TYPE "UDT_Conv_MultiControl_Status"
VERSION : 0.1
   STRUCT
      OL_Maintenance_Mode : Bool;   // Maintenance mode on
      ER_PE1_Blockage : Bool;   // PE1 blockage
      ER_PE2_Blockage : Bool;   // PE2 blockage
      ER_Motor_1_Fault : Bool;   // Motor has error
      ER_Motor_2_Fault : Bool;   // Motor has error
      ER_Motor_3_Fault : Bool;   // Motor has error
      ER_Motor_4_Fault : Bool;   // Motor has error
      ER_Motor_5_Fault : Bool;   // Motor has error
      ER_Motor_6_Fault : Bool;   // Motor has error
      ER_Motor_7_Fault : Bool;   // Motor has error
      ER_Motor_8_Fault : Bool;   // Motor has error
      ER_Motor_9_Fault : Bool;   // Motor has error
      ER_Motor_10_Fault : Bool;   // Motor has error
      ER_Motor_11_Fault : Bool;   // Motor has error
      ER_Motor_12_Fault : Bool;   // Motor has error
      ER_Motor_13_Fault : Bool;   // Motor has error
      ER_Motor_14_Fault : Bool;   // Motor has error
      ER_Motor_15_Fault : Bool;   // Motor has error
      ER_Motor_16_Fault : Bool;   // Motor has error
      Spare_2_3 : Bool;   // Spare_2_3
      Spare_2_4 : Bool;   // Spare_2_4
      Spare_2_5 : Bool;   // Spare_2_5
      Spare_2_6 : Bool;   // Spare_2_6
      Spare_2_7 : Bool;   // Spare_2_7
      Spare_3_0 : Bool;   // Spare_3_0
      Spare_3_1 : Bool;   // Spare_3_1
      Spare_3_2 : Bool;   // Spare_3_2
      Spare_3_3 : Bool;   // Spare_3_3
      Spare_3_4 : Bool;   // Spare_3_4
      Spare_3_5 : Bool;   // Spare_3_5
      Spare_3_6 : Bool;   // Spare_3_6
      Spare_3_7 : Bool;   // Spare_3_7
   END_STRUCT;

END_TYPE

FUNCTION_BLOCK "FB_HW_VFD_G115D"
{ S7_Optimized_Access := 'TRUE' }
VERSION : 0.1
   VAR_INPUT
      i_Telegram_HW_ID { ExternalAccessible := 'False'; ExternalVisible := 'False'; ExternalWritable := 'False'} : HW_SUBMODULE;
      i_Additional_HW_ID { ExternalAccessible := 'False'; ExternalVisible := 'False'; ExternalWritable := 'False'} : HW_SUBMODULE;
      i_Enable : Bool;
      i_IO_Available : Bool;
      i_Safety_OK : Bool := TRUE;
      i_CMD_Reset : Bool;
      i_CMD_Clear_Stat : Bool;
      i_HW_Setting : "UDT_G115D_Setting";
      i_CFG_Motor_Switch_Time : Int := 500;
      i_CMD_Select_Speed : Int := 1;
      i_CMD_Motor_Run : Bool;
      i_CMD_Motor_Reverse : Bool;
   END_VAR

   VAR_OUTPUT RETAIN
      o_Ready_To_Reset : Bool;
      o_Req_Halt : Bool;
      o_ER_PN_Not_Present : Bool;
      o_ER_PN_Error : Bool;
      o_ER_Motor_Fault : Bool;
      o_WN_Motor_Alarm : Bool;
      o_ER_STO_Active : Bool;
      o_WN_No_MemoryCard : Bool;
      o_ST_Motor_Running : Bool;
      o_FaultCode : Word;
      o_AlarmCode : Word;
      o_Speed_Selected : Int;
   END_VAR
   VAR_OUTPUT
      o_Diagnostics : "UDT_G115D_HW_Diagnostics";
   END_VAR

   VAR_IN_OUT
      io_Global : "UDT_Global";
      io_G115D_Interface : "UDT_G115D_HW_Interface";
   END_VAR

   VAR
      s_FB_SINA_SPEED_TEL1 { S7_SetPoint := 'False'} : "FB_SINA_SPEED_TEL1";
   END_VAR
   VAR RETAIN
      s_Copy : Struct
         Clear_Stat : Bool;
         MTR_Run : Bool;
         MTR_Reverse : Bool;
      END_STRUCT;
      s_Motor_Switch_Action_Delay : Int;
      s_Timer_Reset_Delay : Int;
      s_HW_ConfigAxis : Word := 16#003F;
      s_HW_Actual_Speed : Int;
      s_Motor_Run : Bool;
      s_Switch_In_Progress : Bool;
      s_Stopped_Elapsed : Bool;
      s_CMD_Reset : Bool;
      s_HW_Enabled : Bool;
      s_HW_Lockout : Bool;
      s_HW_Fault : Bool;
      s_HW_Alarm : Bool;
   END_VAR

   VAR_TEMP
      t_GeoAddr {InstructionName := 'GEOADDR'; LibVersion := '1.0'} : GEOADDR;
      t_Ret_Val_Int : Int;
      t_Start_Address : Int;
      t_Speed_Setpoint : Int;
      t_IO_Available : Bool;
      t_Enable_Axis : Bool;
   END_VAR

   VAR CONSTANT
      C_RESET_DELAY_TIME : Int := 200;
   END_VAR


BEGIN
	REGION NETOWRK: Initial
	    #o_Ready_To_Reset := FALSE;
	END_REGION

	REGION NETOWRK: Diagnose PN Status
	    #t_Ret_Val_Int := LOG2GEO(LADDR := #i_Telegram_HW_ID, GEOADDR := #t_GeoAddr);
	    IF #i_CMD_Reset OR NOT #i_IO_Available THEN
	        #o_ER_PN_Not_Present := FALSE;
	        #o_ER_PN_Error := FALSE;
	    END_IF;
	    IF #i_IO_Available AND (#t_Ret_Val_Int <> 0 OR "DB_Diagnostics".PNIO_System_100.Device_Not_Present[#t_GeoAddr.STATION]) THEN
	        #o_ER_PN_Not_Present := TRUE;
	    END_IF;
	    IF #i_IO_Available AND "DB_Diagnostics".PNIO_System_100.Device_Error[#t_GeoAddr.STATION] THEN
	        #o_ER_PN_Error := TRUE;
	    END_IF;
	    IF
	        #o_ER_PN_Not_Present AND NOT (#t_Ret_Val_Int <> 0 OR "DB_Diagnostics".PNIO_System_100.Device_Not_Present[#t_GeoAddr.STATION])
	        //OR (#o_ER_PN_Error AND NOT "DB_Diagnostics".PNIO_System_100.Device_Error[#t_GeoAddr.STATION])
	    THEN
	        #o_Ready_To_Reset := TRUE;
	    END_IF;
	    #t_IO_Available := #i_IO_Available AND NOT #o_ER_PN_Not_Present;
	END_REGION

	REGION NETWORK: Read IO
	    "FC_IFM_VFD_G115D_In"(i_Telegram_HW_ID            := #i_Telegram_HW_ID,
	                          i_Additional_HW_ID          := #i_Additional_HW_ID,
	                          o_Telegram_Start_Address    => #t_Start_Address,
	                          o_ActualValue_Start_Address => #t_Start_Address,
	                          o_Data                      => #io_G115D_Interface.Input);
	END_REGION

	REGION NETOWRK: Motor switch delay
	    IF #i_CMD_Motor_Reverse XOR #s_Copy.MTR_Reverse THEN
	        #s_Switch_In_Progress := TRUE;
	        #o_Diagnostics.Motor_Direction_Switch_Count += 1;
	    END_IF;

	    "FC_Delay_On"(i_CMD_Start     := #s_Motor_Run,
	                  i_CFG_Target    := #i_CFG_Motor_Switch_Time,
	                  i_Cycle_Count   := #io_Global.OB_Prev_Cycle_Time,
	                  o_Delay_Finish => #s_Stopped_Elapsed,
	                  io_Setpoint     := #s_Motor_Switch_Action_Delay);

	    IF NOT #s_Stopped_Elapsed THEN
	        #s_Switch_In_Progress := FALSE;
	    END_IF;
	    #o_Req_Halt := #s_Switch_In_Progress;
	END_REGION

	REGION NETOWRK: Reset Pulse
	    "FC_Delay_Off"(i_CMD_Start     := #i_CMD_Reset AND #t_IO_Available,
	                   i_CFG_Target    := #C_RESET_DELAY_TIME,
	                   i_Cycle_Count   := #io_Global.OB_Prev_Cycle_Time,
	                   o_Delay_Finish => #s_CMD_Reset,
	                   io_Setpoint     := #s_Timer_Reset_Delay);
	END_REGION

	REGION NETOWRK: Choose Speedsetpoint
	    IF #i_CMD_Select_Speed = 0 THEN
	        #o_Speed_Selected := #i_HW_Setting.Speed1;
	    ELSIF #i_CMD_Select_Speed = 1 THEN
	        #o_Speed_Selected := #i_HW_Setting.Speed2;
	    ELSIF #i_CMD_Select_Speed = 2 THEN
	        #o_Speed_Selected := #i_HW_Setting.Speed3;
	    ELSIF #i_CMD_Select_Speed = 3 THEN
	        #o_Speed_Selected := #i_HW_Setting.Speed4;
	    ELSE
	        #o_Speed_Selected := #i_HW_Setting.Speed1;
	    END_IF;
	END_REGION

	REGION NETOWRK: 1# Telegram
	    #s_Motor_Run := #i_CMD_Motor_Run AND #t_IO_Available AND NOT #o_ER_Motor_Fault AND NOT #o_ER_STO_Active AND NOT #s_Switch_In_Progress;

	    #s_HW_ConfigAxis := 16#003F;
	    #s_HW_ConfigAxis.%X3 := #i_Safety_OK;
	    #s_HW_ConfigAxis.%X6 := #i_HW_Setting.ReverseDirection XOR #i_CMD_Motor_Reverse;

	    IF #i_HW_Setting.Magnetization_Delay <= 0 THEN
	        IF #s_Motor_Run THEN
	            #t_Speed_Setpoint := #o_Speed_Selected;
	        ELSE
	            #t_Speed_Setpoint := 0;
	        END_IF;
	        #t_Enable_Axis := #i_Enable AND NOT #o_ER_Motor_Fault AND NOT #o_ER_STO_Active;
	    ELSE
	        #t_Enable_Axis := #s_Motor_Run;
	        #t_Speed_Setpoint := #o_Speed_Selected;
	    END_IF;

	    #s_FB_SINA_SPEED_TEL1(EnableAxis      := #t_Enable_Axis,
	                          AckError        := #s_CMD_Reset,
	                          SpeedSetpoint   := #t_Speed_Setpoint,
	                          RefSpeed        := #i_HW_Setting.RefSpeed,
	                          Acceleration    := #i_HW_Setting.Acceleration,
	                          Deceleration    := #i_HW_Setting.Deceleration,
	                          RefRampTime     := #i_HW_Setting.RefRampTime,
	                          ConfigAxis      := #s_HW_ConfigAxis,
	                          AxisEnabled     => #s_HW_Enabled,
	                          Lockout         => #s_HW_Lockout,
	                          Fault           => #s_HW_Fault,
	                          Alarm           => #s_HW_Alarm,
	                          ActualSpeed     => #s_HW_Actual_Speed,
	                          FaultCode       => #o_FaultCode,
	                          AlarmCode       => #o_AlarmCode,
	                          io_HW_Interface := #io_G115D_Interface);
	END_REGION

	REGION NETOWRK: Motor Status
	    #o_ST_Motor_Running := #t_Enable_Axis AND #s_HW_Actual_Speed <> 0;

	    IF #s_CMD_Reset OR NOT #t_IO_Available OR NOT #i_Safety_OK THEN
	        #o_ER_Motor_Fault := FALSE;
	        #o_ER_STO_Active := FALSE;
	    END_IF;

	    IF #t_IO_Available AND #i_Safety_OK AND (#s_HW_Fault OR #s_HW_Lockout) THEN
	        #o_ER_Motor_Fault := TRUE;
	    END_IF;

	    IF #o_ER_Motor_Fault AND NOT (#s_HW_Fault OR #s_HW_Lockout) THEN
	        #o_Ready_To_Reset := TRUE;
	    END_IF;

	    #o_WN_Motor_Alarm :=  #t_IO_Available AND #i_Safety_OK AND #s_HW_Alarm;
	    #o_WN_No_MemoryCard := #t_IO_Available AND NOT #io_G115D_Interface.Input.ZSW2_G115D_Bit00_Memory_Card_In;

	    IF
	        #t_IO_Available
	        AND #i_Safety_OK
	        AND #i_HW_Setting.STOUsed
	        AND (NOT #io_G115D_Interface.Input.ZSW_G115D_Bit02_DI2
	        OR NOT #io_G115D_Interface.Input.ZSW_G115D_Bit03_DI3
	        OR #io_G115D_Interface.Input.ZSW_G115D_Bit06_STOActive)
	    THEN
	        #o_ER_STO_Active := TRUE;
	    END_IF;

	    IF
	        #o_ER_STO_Active
	        AND NOT (NOT #io_G115D_Interface.Input.ZSW_G115D_Bit02_DI2
	        OR NOT #io_G115D_Interface.Input.ZSW_G115D_Bit03_DI3
	        OR #io_G115D_Interface.Input.ZSW_G115D_Bit06_STOActive)
	    THEN
	        #o_Ready_To_Reset := TRUE;
	    END_IF;
	END_REGION

	REGION NETWORK: Write IO
	    "FC_IFM_VFD_G115D_Out"(i_Telegram_HW_ID            := #i_Telegram_HW_ID,
	                           i_Additional_HW_ID          := #i_Additional_HW_ID,
	                           i_Data                      := #io_G115D_Interface.Output,
	                           o_Telegram_Start_Address    => #t_Start_Address,
	                           o_ActualValue_Start_Address => #t_Start_Address);
	END_REGION

	REGION NETOWRK: Diagnostics and Statistical
	    #o_Diagnostics.Run_Command := #t_Enable_Axis AND #t_Speed_Setpoint <> 0;
	    #o_Diagnostics.Brake_Open := #io_G115D_Interface.Input.ZSW1_Bit12_Brake;
	    #o_Diagnostics.DI0 := #io_G115D_Interface.Input.ZSW_G115D_Bit00_DI0;
	    #o_Diagnostics.DI1 := #io_G115D_Interface.Input.ZSW_G115D_Bit01_DI1;
	    #o_Diagnostics.DI2 := #io_G115D_Interface.Input.ZSW_G115D_Bit02_DI2;
	    #o_Diagnostics.DI3 := #io_G115D_Interface.Input.ZSW_G115D_Bit03_DI3;
	    #o_Diagnostics.DIO24 := #io_G115D_Interface.Input.ZSW_G115D_Bit04_DIO24 OR #io_G115D_Interface.Output.STW_G115D_Bit00_DO24;
	    #o_Diagnostics.DIO25 := #io_G115D_Interface.Input.ZSW_G115D_Bit05_DIO25 OR #io_G115D_Interface.Output.STW_G115D_Bit01_DO25;
	    #o_Diagnostics.Memory_Card_In := #io_G115D_Interface.Input.ZSW2_G115D_Bit00_Memory_Card_In;
	    #o_Diagnostics.Memory_Card_Active := #io_G115D_Interface.Input.ZSW2_G115D_Bit01_Memory_Card_Active;
	    #o_Diagnostics.PN_Port1_Down := FALSE;
	    #o_Diagnostics.PN_Port2_Down := FALSE;
	    #o_Diagnostics.Actual_Speed := #s_HW_Actual_Speed;
	    #o_Diagnostics.DCLink_Voltage := #io_G115D_Interface.Input.DCLinkVoltage;
	    #o_Diagnostics.Actual_Current := #io_G115D_Interface.Input.ActualCurrent;
	    #o_Diagnostics.Active_Power := #io_G115D_Interface.Input.ActivePower;

	    IF #o_ST_Motor_Running AND NOT #s_Copy.MTR_Run THEN
	        #o_Diagnostics.Motor_Start_Stop_Count += 1;
	    END_IF;

	    IF #o_ST_Motor_Running AND #io_Global.OS_New_Second THEN
	        #o_Diagnostics.Motor_Started_Time += 1;
	    END_IF;

	    IF #i_CMD_Clear_Stat AND NOT #s_Copy.Clear_Stat THEN
	        #o_Diagnostics.Motor_Started_Time := 0;
	        #o_Diagnostics.Motor_Start_Stop_Count := 0;
	        #o_Diagnostics.Motor_Direction_Switch_Count := 0;
	    END_IF;
	END_REGION

	REGION NETOWRK: Storage Previous State
	    #s_Copy.MTR_Run := #o_ST_Motor_Running;
	    #s_Copy.MTR_Reverse := #i_CMD_Motor_Reverse;
	    #s_Copy.Clear_Stat := #i_CMD_Clear_Stat;
	END_REGION

END_FUNCTION_BLOCK

TYPE "UDT_Conv_G115D_Status"
VERSION : 0.1
   STRUCT
      OL_Maintenance_Mode : Bool;   // Maintenance mode on
      ER_PE1_Blockage : Bool;   // PE1 blockage
      ER_PE2_Blockage : Bool;   // PE2 blockage
      ER_VFD_PN_NotPresent : Bool;   // VFD not present on profinet network
      ER_VFD_PN_Error : Bool;   // VFD has error profinet network
      ER_VFD_Fault : Bool;   // VFD has error
      WN_VFD_Alarm : Bool;   // VFD has an warning
      ER_VFD_STO_Active : Bool;   // VFD STO is active
      WN_No_MemoryCard : Bool;   // Memory card is missing
      Spare_1_1 : Bool;   // Spare_1_1
      Spare_1_2 : Bool;   // Spare_1_2
      Spare_1_3 : Bool;   // Spare_1_3
      Spare_1_4 : Bool;   // Spare_1_4
      Spare_1_5 : Bool;   // Spare_1_5
      Spare_1_6 : Bool;   // Spare_1_6
      Spare_1_7 : Bool;   // Spare_1_7
      FaultCode : Word;   // VFD fault code
      AlarmCode : Word;   // VFD alarm code
   END_STRUCT;

END_TYPE

TYPE "UDT_Conv_G115D_Command"
VERSION : 0.1
   STRUCT
      Man_Mode : Bool;   // Maintenance mode on
      Man_Clear : Bool;   // Maintenance - Clear data
      Man_Run : Bool;   // Maintenance - Run motor
      Man_DisableAxis : Bool;   // Maintenance - Disable axis
      Cmd_Reset_ESave : Bool;   // Command - Reset energy save
      Cmd_Bypass_Fault : Bool;   // Command - Bypass all fault
      Spare_0_6 : Bool;   // Spare_0_6
      Spare_0_7 : Bool;   // Spare_0_7
      Spare_1_0 : Bool;   // Spare_1_0
      Spare_1_1 : Bool;   // Spare_1_1
      Spare_1_2 : Bool;   // Spare_1_2
      Spare_1_3 : Bool;   // Spare_1_3
      Spare_1_4 : Bool;   // Spare_1_4
      Spare_1_5 : Bool;   // Spare_1_5
      Spare_1_6 : Bool;   // Spare_1_6
      Spare_1_7 : Bool;   // Spare_1_7
   END_STRUCT;

END_TYPE

TYPE "UDT_PAC_HW_Input"
VERSION : 0.1
   STRUCT
      Status_Bit00_SynchronizationMissing : Bool;
      Status_Bit01_ConfigurationMenuActive : Bool;
      Status_Bit02_VoltageOverload : Bool;
      Status_Bit03_CurrentOverload : Bool;
      Status_Bit04_Reserved : Bool;
      Status_Bit05_Reserved : Bool;
      Status_Bit06_WriteProtectionActive : Bool;
      Status_Bit07_Reserved : Bool;
      Status_Bit08_Reserved : Bool;
      Status_Bit09_MaximumPulseRateExceeded : Bool;
      Status_Bit10_Reserved : Bool;
      Status_Bit11_Reserved : Bool;
      Status_Bit12_Reserved : Bool;
      Status_Bit13_Reserved : Bool;
      Status_Bit14_Reserved : Bool;
      Status_Bit15_Reserved : Bool;
      Status_Bit16_ConfigurationChanged : Bool;
      Status_Bit17_LimitViolation : Bool;
      Status_Bit18_PulseRateExceededStored : Bool;
      Status_Bit19_Reserved : Bool;
      Status_Bit20_Reserved : Bool;
      Status_Bit21_Reserved : Bool;
      Status_Bit22_Reserved : Bool;
      Status_Bit23_Reserved : Bool;
      Status_Bit24_Reserved : Bool;
      Status_Bit25_Reserved : Bool;
      Status_Bit26_Reserved : Bool;
      Status_Bit27_Reserved : Bool;
      Status_Bit28_Reserved : Bool;
      Status_Bit29_Reserved : Bool;
      Status_Bit30_Reserved : Bool;
      Status_Bit31_Reserved : Bool;
      Voltage_L1_N : Real;
      Voltage_L2_N : Real;
      Voltage_L3_N : Real;
      Voltage_L1_L2 : Real;
      Voltage_L2_L3 : Real;
      Voltage_L3_L1 : Real;
      Current_L1 : Real;
      Current_L2 : Real;
      Current_L3 : Real;
      PowerFactor_L1 : Real;
      PowerFactor_L2 : Real;
      PowerFactor_L3 : Real;
      THD_Voltage_L1 : Real;
      THD_Voltage_L2 : Real;
      THD_Voltage_L3 : Real;
      THD_Current_L1 : Real;
      THD_Current_L2 : Real;
      THD_Current_L3 : Real;
      Frequency : Real;
      Average_Current : Real;
      Total_ApparentPower : Real;
      Total_ActivePower : Real;
      Total_ReactivePower : Real;
      Total_PowerFactor : Real;
      Amplitude_Unbalance_Voltage : Real;
      Amplitude_Unbalance_Current : Real;
      Last_Period_Length : Real;
   END_STRUCT;

END_TYPE

TYPE "UDT_PAC_HW_Output"
VERSION : 0.1
   STRUCT
      Control_Bit00_ResetMaximumValues : Bool;
      Control_Bit01_ResetMinimumValues : Bool;
      Control_Bit02_ResetEnergyCounters : Bool;
      Control_Bit03_AcknowledgeDiagnostics : Bool;
      Control_Bit04_SynchronizeDemandPeriod : Bool;
      Control_Bit05_ProcessCounterStartStop : Bool;
      Control_Bit06_CopyAndResetProcessCounter : Bool;
      Control_Bit07_ResetProcessCounter : Bool;
      Control_Bit08_SwitchHighTariff : Bool;
      Control_Bit09_SwitchLowTariff : Bool;
      Control_Bit10_SwitchOutput00 : Bool;
      Control_Bit11_SwitchOutput01 : Bool;
      Control_Bit12_Reserved : Bool;
      Control_Bit13_Reserved : Bool;
      Control_Bit14_Reserved : Bool;
      Control_Bit15_Reserved : Bool;
   END_STRUCT;

END_TYPE

TYPE "UDT_Accmulation_Command"
VERSION : 0.1
   STRUCT
      Disable : Bool;
      Cleanup : Bool;
   END_STRUCT;

END_TYPE

TYPE "UDT_Conv_Triple_G115D_Command"
VERSION : 0.1
   STRUCT
      Man_Mode : Bool;   // Maintenance mode on
      Man_Clear : Bool;   // Maintenance - Clear data
      Man_Run : Bool;   // Maintenance - Run motor
      Man_DisableAxis : Bool;   // Maintenance - Disable axis
      Cmd_Reset_ESave : Bool;   // Command - Reset energy save
      Cmd_Bypass_Fault : Bool;   // Command - Bypass all fault
      Spare_0_6 : Bool;
      Spare_0_7 : Bool;   // Spare_0_7
      Spare_1_0 : Bool;   // Spare_1_0
      Spare_1_1 : Bool;   // Spare_1_1
      Spare_1_2 : Bool;   // Spare_1_2
      Spare_1_3 : Bool;   // Spare_1_3
      Spare_1_4 : Bool;   // Spare_1_4
      Spare_1_5 : Bool;   // Spare_1_5
      Spare_1_6 : Bool;   // Spare_1_6
      Spare_1_7 : Bool;   // Spare_1_7
   END_STRUCT;

END_TYPE

TYPE "UDT_Ray26_IO"
VERSION : 0.1
   STRUCT
      IsCleared : Bool;
      TechIn : Bool;
      Port_Healthy : Bool;
   END_STRUCT;

END_TYPE

TYPE "UDT_UPS_HW_Input"
VERSION : 0.1
   STRUCT
      Input_Voltage_OK : Bool;
      Buffer_Mode_Active : Bool;
      Ready_For_Buffer : Bool;
      Charge_Sufficient : Bool;
      Need_Change_Battery : Bool;
      Battery_Connection_Fault : Bool;
      Battery_Level : Int;
   END_STRUCT;

END_TYPE

TYPE "UDT_Induct_On_Gap_Command"
VERSION : 0.1
   STRUCT
      Disable_Induct : Bool;
   END_STRUCT;

END_TYPE

TYPE "UDT_Merge_2_To_1_Command"
VERSION : 0.1
   STRUCT
      Disable_Line1 : Bool;
      Disable_Line2 : Bool;
   END_STRUCT;

END_TYPE

TYPE "UDT_IOLink_Master_Command"
VERSION : 0.1
   STRUCT
      CMD_Backup : Bool;
      CMD_Restore : Bool;
      Spare_0_2 : Bool;
      Spare_0_3 : Bool;
      Spare_0_4 : Bool;
      Spare_0_5 : Bool;
      Spare_0_6 : Bool;
      Spare_0_7 : Bool;
      Spare_1_0 : Bool;
      Spare_1_1 : Bool;
      Spare_1_2 : Bool;
      Spare_1_3 : Bool;
      Spare_1_4 : Bool;
      Spare_1_5 : Bool;
      Spare_1_6 : Bool;
      Spare_1_7 : Bool;
      CMD_Trigger_Ray26_Techin : Int;
      CMD_Read_Ray26_Techin_State : Int;
   END_STRUCT;

END_TYPE

TYPE "UDT_Datalogic_AV900_Command"
VERSION : 0.1
   STRUCT
      Cmd_Disable : Bool;
      Spare_0_1 : Bool;
      Spare_0_2 : Bool;
      Spare_0_3 : Bool;
      Spare_0_4 : Bool;
      Spare_0_5 : Bool;
      Spare_0_6 : Bool;
      Spare_0_7 : Bool;
      Spare_1_0 : Bool;
      Spare_1_1 : Bool;
      Spare_1_2 : Bool;
      Spare_1_3 : Bool;
      Spare_1_4 : Bool;
      Spare_1_5 : Bool;
      Spare_1_6 : Bool;
      Spare_1_7 : Bool;
   END_STRUCT;

END_TYPE

TYPE "UDT_ADTA_Command"
VERSION : 0.1
   STRUCT
      Spare_0_0 : Bool;
      Spare_0_1 : Bool;
      Spare_0_2 : Bool;
      Spare_0_3 : Bool;
      Spare_0_4 : Bool;
      Spare_0_5 : Bool;
      Spare_0_6 : Bool;
      Spare_0_7 : Bool;
      Spare_1_0 : Bool;
      Spare_1_1 : Bool;
      Spare_1_2 : Bool;
      Spare_1_3 : Bool;
      Spare_1_4 : Bool;
      Spare_1_5 : Bool;
      Spare_1_6 : Bool;
      Spare_1_7 : Bool;
   END_STRUCT;

END_TYPE

TYPE "UDT_NBS_Command"
VERSION : 0.1
   STRUCT
      Spare_0_0 : Bool;
      Spare_0_1 : Bool;
      Spare_0_2 : Bool;
      Spare_0_3 : Bool;
      Spare_0_4 : Bool;
      Spare_0_5 : Bool;
      Spare_0_6 : Bool;
      Spare_0_7 : Bool;
      Spare_1_0 : Bool;
      Spare_1_1 : Bool;
      Spare_1_2 : Bool;
      Spare_1_3 : Bool;
      Spare_1_4 : Bool;
      Spare_1_5 : Bool;
      Spare_1_6 : Bool;
      Spare_1_7 : Bool;
   END_STRUCT;

END_TYPE

TYPE "UDT_Merge_Singulator_Command"
VERSION : 0.1
   STRUCT
      Spare_0_0 : Bool;
      Spare_0_1 : Bool;
      Spare_0_2 : Bool;
      Spare_0_3 : Bool;
      Spare_0_4 : Bool;
      Spare_0_5 : Bool;
      Spare_0_6 : Bool;
      Spare_0_7 : Bool;
      Spare_1_0 : Bool;
      Spare_1_1 : Bool;
      Spare_1_2 : Bool;
      Spare_1_3 : Bool;
      Spare_1_4 : Bool;
      Spare_1_5 : Bool;
      Spare_1_6 : Bool;
      Spare_1_7 : Bool;
   END_STRUCT;

END_TYPE

TYPE "UDT_Merge_3_To_1_Command"
VERSION : 0.1
   STRUCT
      Disable_Line1 : Bool;
      Disable_Line2 : Bool;
      Disable_Line3 : Bool;
   END_STRUCT;

END_TYPE

TYPE "UDT_SSM_Status"
TITLE = UDT_Status_SSM
VERSION : 0.1
//Status for start stop manager
//# Block Info
//- Title:            UDT_Status_SSM
//- Comment/Function: Status for start stop manager
//- Library/Family:   APS
//- Author:           Jay Liu
//- Tested with:      ---
//- Engineering:      TIA Portal V20
//- Restrictions:     ---
//- Requirements:     ---
//
//# History
// |Version  | Date       | Author                 | Description                   |
// |---------|------------|------------------------|------------------------------ |
// |01.00.00 | 2026-01-22 | Jay Liu                | First released version        |
   STRUCT
      Started : Bool := FALSE;   // Started
      Starting : Bool := FALSE;   // Starting
      Stopped : Bool := FALSE;   // Stopped
      Stopping : Bool := FALSE;   // Stopping
      Ready_To_Restart : Bool := FALSE;   // Ready to restart
      Ready_To_Reset : Bool := FALSE;   // Ready to reset
      Spare_0_6 : Bool := FALSE;   // Spare_0_6
      Spare_0_7 : Bool := FALSE;   // Spare_0_7
      Spare_1_0 : Bool := FALSE;   // Spare_1_0
      Spare_1_1 : Bool := FALSE;   // Spare_1_1
      Spare_1_2 : Bool := FALSE;   // Spare_1_2
      Spare_1_3 : Bool := FALSE;   // Spare_1_3
      Spare_1_4 : Bool := FALSE;   // Spare_1_4
      Spare_1_5 : Bool := FALSE;   // Spare_1_5
      Spare_1_6 : Bool := FALSE;   // Spare_1_6
      Spare_1_7 : Bool := FALSE;   // Spare_1_7
   END_STRUCT;

END_TYPE

TYPE "UDT_SDC_4Servos_Status"
TITLE = UDT_Status_MCC
VERSION : 0.1
//Status of main control cabinet
//# Block Info
//- Title:            UDT_Status_MCC
//- Comment/Function: Status of main control cabinet
//- Library/Family:   APS
//- Author:           Jay Liu
//- Tested with:      ---
//- Engineering:      TIA Portal V20
//- Restrictions:     ---
//- Requirements:     ---
//
//# History
// |Version  | Date       | Author                 | Description                   |
// |---------|------------|------------------------|------------------------------ |
// |01.00.00 | 2026-01-22 | Jay Liu                | First released version        |
   STRUCT
      ER_Main_Switch_Trip : Bool;   // Main switch on cabinet is off
      ER_CB_Q0111_Trip_PowerSupply : Bool;   // Circuit breaker of power supply is off
      ER_Power_Supply_G0111_Fault : Bool;   // 24V Power supply is not ok
      ER_CB_F1002_Trip_Fan : Bool;   // Circuit breaker of fan is off
      WN_Cabinet_Temperature_High : Bool;   // Temperature is high in cabinet
      ER_CB_Q1041_Trip_Servo1 : Bool;   // Motor power of 1# servo is off
      ER_CB_F1041_Trip_Servo1 : Bool;   // Control power of 1# servo is off
      ER_CB_Q1051_Trip_Servo2 : Bool;   // Motor power of 2# servo is off
      ER_CB_F1051_Trip_Servo2 : Bool;   // Control power of 2# servo is off
      ER_CB_Q1061_Trip_Servo3 : Bool;   // Motor power of 3# servo is off
      ER_CB_F1016_Trip_Servo3 : Bool;   // Control power of 3# servo is off
      ER_CB_Q1071_Trip_Servo4 : Bool;   // Motor power of 4# servo is off
      ER_CB_F1071_Trip_Servo4 : Bool;   // Control power of 4# servo is off
      Spare_1_5 : Bool;   // Spare_1_5
      Spare_1_6 : Bool;   // Spare_1_6
      Spare_1_7 : Bool;   // Spare_1_7
      Spare_2_0 : Bool;   // Spare_2_0
      Spare_2_1 : Bool;   // Spare_2_1
      Spare_2_2 : Bool;   // Spare_2_2
      Spare_2_3 : Bool;   // Spare_2_3
      Spare_2_4 : Bool;   // Spare_2_4
      Spare_2_5 : Bool;   // Spare_2_5
      Spare_2_6 : Bool;   // Spare_2_6
      Spare_2_7 : Bool;   // Spare_2_7
      Spare_3_0 : Bool;   // Spare_3_0
      Spare_3_1 : Bool;   // Spare_3_1
      Spare_3_2 : Bool;   // Spare_3_2
      Spare_3_3 : Bool;   // Spare_3_3
      Spare_3_4 : Bool;   // Spare_3_4
      Spare_3_5 : Bool;   // Spare_3_5
      Spare_3_6 : Bool;   // Spare_3_6
      Spare_3_7 : Bool;   // Spare_3_7
   END_STRUCT;

END_TYPE

TYPE "UDT_AC_IO_Status"
TITLE = UDT_Status_MCC
VERSION : 0.1
//Status of main control cabinet
//# Block Info
//- Title:            UDT_Status_MCC
//- Comment/Function: Status of main control cabinet
//- Library/Family:   APS
//- Author:           Jay Liu
//- Tested with:      ---
//- Engineering:      TIA Portal V20
//- Restrictions:     ---
//- Requirements:     ---
//
//# History
// |Version  | Date       | Author                 | Description                   |
// |---------|------------|------------------------|------------------------------ |
// |01.00.00 | 2026-01-22 | Jay Liu                | First released version        |
   STRUCT
      ER_UR20_Not_Present : Bool;   // Profinet module is not present
      ER_UR20_Error : Bool;   // Profinet module has an error
      ER_UPS_Not_Present : Bool;
      ER_UPS_Error : Bool;
      ER_PAC3220_Not_Present : Bool;
      ER_PAC3220_Error : Bool;
      ER_XC208_Not_Present : Bool;
      ER_XC208_Error : Bool;
      ER_XC216_Not_Present : Bool;
      ER_XC216_Error : Bool;
      ER_Breaker_Off_F1062 : Bool;
      ER_Breaker_Off_F1063 : Bool;
      ER_Breaker_Off_F1064 : Bool;
      ER_Breaker_Off_F1065 : Bool;
      ER_Breaker_Off_F1071 : Bool;
      ER_Breaker_Off_F1072 : Bool;
      ER_Breaker_Off_F1073 : Bool;
      ER_Breaker_Off_F1074 : Bool;
      ER_Breaker_Off_F1075 : Bool;
      ER_Breaker_Off_F1151 : Bool;
      ER_Breaker_Off_F1152 : Bool;
      ER_Breaker_Off_F1153 : Bool;
      ER_Breaker_Off_F1161 : Bool;
      ER_Breaker_Off_F1162 : Bool;
      ER_Breaker_Off_F1163 : Bool;
      ER_Breaker_Off_F1171 : Bool;
      ER_Breaker_Off_F1172 : Bool;
      ER_Breaker_Off_F1173 : Bool;
      ER_Breaker_Off_F1181 : Bool;
      ER_Breaker_Off_F1182 : Bool;
      ER_Breaker_Off_F1183 : Bool;
      ER_Breaker_Off_F1191 : Bool;
      ER_Breaker_Off_F1192 : Bool;
      ER_Breaker_Off_F1193 : Bool;
      ER_Breaker_Off_F1501 : Bool;
      ER_Breaker_Off_F1502 : Bool;
      ER_Breaker_Off_F1503 : Bool;
      ER_Breaker_Off_F1504 : Bool;
      ER_Breaker_Off_F1511 : Bool;
      ER_Breaker_Off_F1512 : Bool;
      ER_Breaker_Off_F1513 : Bool;
      ER_Breaker_Off_F1514 : Bool;
      ER_Breaker_Off_F1521 : Bool;
      ER_Breaker_Off_F1522 : Bool;
      ER_Breaker_Off_F1523 : Bool;
      ER_Breaker_Off_F1515 : Bool;
      ER_Breaker_Off_F1516 : Bool;
      ER_Breaker_Off_F1524 : Bool;
      ER_Breaker_Off_F1525 : Bool;
      ER_Breaker_Off_F1526 : Bool;
      ER_Power_Supply_G01_Fault : Bool;
      ER_Cabinet_Temperature_High : Bool;
      Spare_9_1 : Bool;
      Spare_9_2 : Bool;
      Spare_9_3 : Bool;
      Spare_9_4 : Bool;
      Spare_9_5 : Bool;
      Spare_9_6 : Bool;
      Spare_9_7 : Bool;
      Spare_10_0 : Bool;
      Spare_10_1 : Bool;
      Spare_10_2 : Bool;
      Spare_10_3 : Bool;
      Spare_10_4 : Bool;
      Spare_10_5 : Bool;
      Spare_10_6 : Bool;
      Spare_10_7 : Bool;
      Spare_11_0 : Bool;
      Spare_11_1 : Bool;
      Spare_11_2 : Bool;
      Spare_11_3 : Bool;
      Spare_11_4 : Bool;
      Spare_11_5 : Bool;
      Spare_11_6 : Bool;
      Spare_11_7 : Bool;
   END_STRUCT;

END_TYPE

TYPE "UDT_AC_SWS_Status"
TITLE = UDT_Status_MCC
VERSION : 0.1
//Status of main control cabinet
//# Block Info
//- Title:            UDT_Status_MCC
//- Comment/Function: Status of main control cabinet
//- Library/Family:   APS
//- Author:           Jay Liu
//- Tested with:      ---
//- Engineering:      TIA Portal V20
//- Restrictions:     ---
//- Requirements:     ---
//
//# History
// |Version  | Date       | Author                 | Description                   |
// |---------|------------|------------------------|------------------------------ |
// |01.00.00 | 2026-01-22 | Jay Liu                | First released version        |
   STRUCT
      ER_UR20_Not_Present : Bool;   // Profinet module is not present
      ER_UR20_Error : Bool;   // Profinet module has an error
      ER_UPS_Not_Present : Bool;
      ER_UPS_Error : Bool;
      ER_PAC3220_Not_Present : Bool;
      ER_PAC3220_Error : Bool;
      ER_XC208_Not_Present : Bool;
      ER_XC208_Error : Bool;
      ER_XC216_Not_Present : Bool;
      ER_XC216_Error : Bool;
      ER_Breaker_Off_F1062 : Bool;   // Emergency stop is active
      ER_Breaker_Off_F1063 : Bool;   // External emergency stop is active
      ER_Breaker_Off_F1064 : Bool;   // Spare_1_1
      ER_Breaker_Off_F1065 : Bool;   // Spare_1_2
      ER_Breaker_Off_F1071 : Bool;   // Spare_1_3
      ER_Breaker_Off_F1072 : Bool;   // Spare_1_4
      ER_Breaker_Off_F1073 : Bool;   // Spare_1_5
      ER_Breaker_Off_F1074 : Bool;   // Spare_1_6
      ER_Breaker_Off_F1075 : Bool;   // Spare_1_7
      ER_Breaker_Off_F1151 : Bool;
      ER_Breaker_Off_F1152 : Bool;
      ER_Breaker_Off_F1153 : Bool;
      ER_Breaker_Off_F1161 : Bool;
      ER_Breaker_Off_F1162 : Bool;
      ER_Breaker_Off_F1163 : Bool;
      ER_Breaker_Off_F1171 : Bool;
      ER_Breaker_Off_F1172 : Bool;
      ER_Breaker_Off_F1173 : Bool;
      ER_Breaker_Off_F1181 : Bool;
      ER_Breaker_Off_F1182 : Bool;
      ER_Breaker_Off_F1183 : Bool;
      ER_Breaker_Off_F1191 : Bool;
      ER_Breaker_Off_F1192 : Bool;
      ER_Breaker_Off_F1193 : Bool;
      ER_Breaker_Off_F1501 : Bool;
      ER_Breaker_Off_F1502 : Bool;
      ER_Breaker_Off_F1503 : Bool;
      ER_Breaker_Off_F1504 : Bool;
      ER_Breaker_Off_F1511 : Bool;
      ER_Breaker_Off_F1512 : Bool;
      ER_Breaker_Off_F1513 : Bool;
      ER_Breaker_Off_F1514 : Bool;
      ER_Breaker_Off_F1521 : Bool;
      ER_Breaker_Off_F1522 : Bool;
      ER_Breaker_Off_F1523 : Bool;
      ER_Breaker_Off_F1515 : Bool;
      ER_Breaker_Off_F1516 : Bool;
      ER_Breaker_Off_F1524 : Bool;
      ER_Breaker_Off_F1525 : Bool;
      ER_Breaker_Off_F1526 : Bool;
      ER_Power_Supply_G01_Fault : Bool;
      ER_Cabinet_Temperature_High : Bool;
      Spare_9_1 : Bool;
      Spare_9_2 : Bool;
      Spare_9_3 : Bool;
      Spare_9_4 : Bool;
      Spare_9_5 : Bool;
      Spare_9_6 : Bool;
      Spare_9_7 : Bool;
      Spare_10_0 : Bool;
      Spare_10_1 : Bool;
      Spare_10_2 : Bool;
      Spare_10_3 : Bool;
      Spare_10_4 : Bool;
      Spare_10_5 : Bool;
      Spare_10_6 : Bool;
      Spare_10_7 : Bool;
      Spare_11_0 : Bool;
      Spare_11_1 : Bool;
      Spare_11_2 : Bool;
      Spare_11_3 : Bool;
      Spare_11_4 : Bool;
      Spare_11_5 : Bool;
      Spare_11_6 : Bool;
      Spare_11_7 : Bool;
   END_STRUCT;

END_TYPE

TYPE "UDT_RLS_Command"
VERSION : 0.1
   STRUCT
      Spare_0_0 : Bool;
      Spare_0_1 : Bool;
      Spare_0_2 : Bool;
      Spare_0_3 : Bool;
      Spare_0_4 : Bool;
      Spare_0_5 : Bool;
      Spare_0_6 : Bool;
      Spare_0_7 : Bool;
      Spare_1_0 : Bool;
      Spare_1_1 : Bool;
      Spare_1_2 : Bool;
      Spare_1_3 : Bool;
      Spare_1_4 : Bool;
      Spare_1_5 : Bool;
      Spare_1_6 : Bool;
      Spare_1_7 : Bool;
   END_STRUCT;

END_TYPE

TYPE "UDT_SDC_10Servos_Status"
TITLE = UDT_Status_MCC
VERSION : 0.1
//Status of main control cabinet
//# Block Info
//- Title:            UDT_Status_MCC
//- Comment/Function: Status of main control cabinet
//- Library/Family:   APS
//- Author:           Jay Liu
//- Tested with:      ---
//- Engineering:      TIA Portal V20
//- Restrictions:     ---
//- Requirements:     ---
//
//# History
// |Version  | Date       | Author                 | Description                   |
// |---------|------------|------------------------|------------------------------ |
// |01.00.00 | 2026-01-22 | Jay Liu                | First released version        |
   STRUCT
      ER_Main_Switch_Trip : Bool;   // Main switch on cabinet is off
      ER_CB_Q0111_Trip_Power_Supply : Bool;   // Circuit breaker of power supply is off
      ER_Power_Supply_G0111_Fault : Bool;   // 24V Power supply is not ok
      ER_CB_F1002_Trip_Fan : Bool;   // Circuit breaker of fan is off
      WN_Cabinet_Temperature_High : Bool;   // Temperature is high in cabinet
      ER_CB_Q0401_Trip_Servo1 : Bool;   // Motor power of 1# servo is off
      ER_CB_F0401_Trip_Servo1 : Bool;   // Control power of 1# servo is off
      ER_CB_Q0411_Trip_Servo2 : Bool;   // Motor power of 2# servo is off
      ER_CB_F0411_Trip_Servo2 : Bool;   // Control power of 2# servo is off
      ER_CB_Q0421_Trip_Servo3 : Bool;   // Motor power of 3# servo is off
      ER_CB_F0421_Trip_Servo3 : Bool;   // Control power of 3# servo is off
      ER_CB_Q0431_Trip_Servo4 : Bool;   // Motor power of 4# servo is off
      ER_CB_F0431_Trip_Servo4 : Bool;   // Control power of 4# servo is off
      ER_CB_Q0441_Trip_Servo5 : Bool;   // Motor power of 5# servo is off
      ER_CB_F0441_Trip_Servo5 : Bool;   // Control power of 5# servo is off
      ER_CB_Q0451_Trip_Servo6 : Bool;   // Motor power of 6# servo is off
      ER_CB_F0451_Trip_Servo6 : Bool;   // Control power of 6# servo is off
      ER_CB_Q0461_Trip_Servo7 : Bool;   // Motor power of 7# servo is off
      ER_CB_F0461_Trip_Servo7 : Bool;   // Control power of 7# servo is off
      ER_CB_Q0471_Trip_Servo8 : Bool;   // Motor power of 8# servo is off
      ER_CB_F0471_Trip_Servo8 : Bool;   // Control power of 8# servo is off
      ER_CB_Q0481_Trip_Servo9 : Bool;   // Motor power of 9# servo is off
      ER_CB_F0481_Trip_Servo9 : Bool;   // Control power of 9# servo is off
      ER_CB_Q0491_Trip_Servo10 : Bool;   // Motor power of 10# servo is off
      ER_CB_F0491_Trip_Servo10 : Bool;   // Control power of 10# servo is off
      Spare_3_1 : Bool;   // Spare_3_1
      Spare_3_2 : Bool;   // Spare_3_2
      Spare_3_3 : Bool;   // Spare_3_3
      Spare_3_4 : Bool;   // Spare_3_4
      Spare_3_5 : Bool;   // Spare_3_5
      Spare_3_6 : Bool;   // Spare_3_6
      Spare_3_7 : Bool;   // Spare_3_7
   END_STRUCT;

END_TYPE

TYPE "UDT_Datalogic_AV900_Status"
VERSION : 0.1
   STRUCT
      ER_PN_NotPresent : Bool;
      ER_PN_Error : Bool;
      OL_Disabled : Bool;
      WN_NoCode : Bool;
      WN_NoRead : Bool;
      WN_MultiRead : Bool;
      WN_InvalidData : Bool;
      WN_UnexpectedData : Bool;
      ER_Successive_NoCode : Bool;
      ER_Successive_NoRead : Bool;
      ER_Successive_MultiRead : Bool;
      ER_Successive_InvalidData : Bool;
      ER_Successive_UnexpectedData : Bool;
      Spare_1_5 : Bool;
      Spare_1_6 : Bool;
      Spare_1_7 : Bool;
      Spare_2_0 : Bool;
   END_STRUCT;

END_TYPE

TYPE "UDT_Tipper_Status"
VERSION : 0.1
   STRUCT
      Spare_0_0 : Bool;
      Spare_0_1 : Bool;
      Spare_0_2 : Bool;
      Spare_0_3 : Bool;
      Spare_0_4 : Bool;
      Spare_0_5 : Bool;
      Spare_0_6 : Bool;
      Spare_0_7 : Bool;
      Spare_1_0 : Bool;
      Spare_1_1 : Bool;
      Spare_1_2 : Bool;
      Spare_1_3 : Bool;
      Spare_1_4 : Bool;
      Spare_1_5 : Bool;
      Spare_1_6 : Bool;
      Spare_1_7 : Bool;
   END_STRUCT;

END_TYPE

TYPE "UDT_Echelon_Status"
VERSION : 0.1
   STRUCT
      ER_PN_NotPresent : Bool;
      ER_PN_Error : Bool;
      Spare_0_2 : Bool;
      Spare_0_3 : Bool;
      Spare_0_4 : Bool;
      Spare_0_5 : Bool;
      Spare_0_6 : Bool;
      Spare_0_7 : Bool;
      Spare_1_0 : Bool;
      Spare_1_1 : Bool;
      Spare_1_2 : Bool;
      Spare_1_3 : Bool;
      Spare_1_4 : Bool;
      Spare_1_5 : Bool;
      Spare_1_6 : Bool;
      Spare_1_7 : Bool;
   END_STRUCT;

END_TYPE

TYPE "UDT_RLS_Status"
VERSION : 0.1
   STRUCT
      ER_PN_NotPresent : Bool;
      ER_PN_Error : Bool;
      Spare_0_2 : Bool;
      Spare_0_3 : Bool;
      Spare_0_4 : Bool;
      Spare_0_5 : Bool;
      Spare_0_6 : Bool;
      Spare_0_7 : Bool;
      Spare_1_0 : Bool;
      Spare_1_1 : Bool;
      Spare_1_2 : Bool;
      Spare_1_3 : Bool;
      Spare_1_4 : Bool;
      Spare_1_5 : Bool;
      Spare_1_6 : Bool;
      Spare_1_7 : Bool;
   END_STRUCT;

END_TYPE

TYPE "UDT_Merge_Singulator_Status"
VERSION : 0.1
   STRUCT
      ER_PN_NotPresent : Bool;
      ER_PN_Error : Bool;
      OL_PassThrough_Mode : Bool;
      OL_Manual_Mode : Bool;
      WN_LowCapacity_Mode : Bool;
      ER_Device_Fault : Bool;
      ER_Jam : Bool;
      ER_Singulate_Ratio_Low : Bool;
      WN_Singulate_Ratio_Low : Bool;
      Spare_1_1 : Bool;
      Spare_1_2 : Bool;
      Spare_1_3 : Bool;
      Spare_1_4 : Bool;
      Spare_1_5 : Bool;
      Spare_1_6 : Bool;
      Spare_1_7 : Bool;
   END_STRUCT;

END_TYPE

TYPE "UDT_NBS_Status"
VERSION : 0.1
   STRUCT
      ER_PN_NotPresent : Bool;
      ER_PN_Error : Bool;
      ER_Communication_Fault : Bool;
      WN_Slow_Mode : Bool;
      OL_PassThrough_Mode : Bool;
      Spare_0_5 : Bool;
      Spare_0_6 : Bool;
      Spare_0_7 : Bool;
      Spare_1_0 : Bool;
      Spare_1_1 : Bool;
      Spare_1_2 : Bool;
      Spare_1_3 : Bool;
      Spare_1_4 : Bool;
      Spare_1_5 : Bool;
      Spare_1_6 : Bool;
      Spare_1_7 : Bool;
   END_STRUCT;

END_TYPE

TYPE "UDT_ADTA_Status"
VERSION : 0.1
   STRUCT
      ER_PN_NotPresent : Bool;
      ER_PN_Error : Bool;
      Spare_0_2 : Bool;
      Spare_0_3 : Bool;
      Spare_0_4 : Bool;
      Spare_0_5 : Bool;
      Spare_0_6 : Bool;
      Spare_0_7 : Bool;
      Spare_1_0 : Bool;
      Spare_1_1 : Bool;
      Spare_1_2 : Bool;
      Spare_1_3 : Bool;
      Spare_1_4 : Bool;
      Spare_1_5 : Bool;
      Spare_1_6 : Bool;
      Spare_1_7 : Bool;
   END_STRUCT;

END_TYPE

TYPE "UDT_IOLink_Master_Status"
VERSION : 0.1
   STRUCT
      ER_PN_NotPresent : Bool;
      ER_PN_Error : Bool;
      ER_Port1_NotHealthy : Bool;
      ER_Port2_NotHealthy : Bool;
      ER_Port3_NotHealthy : Bool;
      ER_Port4_NotHealthy : Bool;
      ER_Port5_NotHealthy : Bool;
      ER_Port6_NotHealthy : Bool;
      ER_Port7_NotHealthy : Bool;
      ER_Port8_NotHealthy : Bool;
      ST_Backup_Data_Valid : Bool;
      WN_Backup_Fault : Bool;
      ST_Restore_Success : Bool;
      WN_Restore_Fault : Bool;
      ST_Port_Command_Success : Bool;
      WN_Port_Command_Fault : Bool;
      Spare_2_0 : Bool;
      Spare_2_1 : Bool;
      Spare_2_2 : Bool;
      Spare_2_3 : Bool;
      Spare_2_4 : Bool;
      Spare_2_5 : Bool;
      Spare_2_6 : Bool;
      Spare_2_7 : Bool;
      Spare_3_0 : Bool;
      Spare_3_1 : Bool;
      Spare_3_2 : Bool;
      Spare_3_3 : Bool;
      Spare_3_4 : Bool;
      Spare_3_5 : Bool;
      Spare_3_6 : Bool;
      Spare_3_7 : Bool;
   END_STRUCT;

END_TYPE

TYPE "UDT_MultiControl_Status"
VERSION : 0.1
   STRUCT
      ER_PN_NotPresent : Bool;
      ER_PN_Error : Bool;
      ER_Motor_Voltage_Fault : Bool;
      WN_Over_Temperature : Bool;
      Spare_0_4 : Bool;
      Spare_0_5 : Bool;
      Spare_0_6 : Bool;
      Spare_0_7 : Bool;
      Spare_1_0 : Bool;
      Spare_1_1 : Bool;
      Spare_1_2 : Bool;
      Spare_1_3 : Bool;
      Spare_1_4 : Bool;
      Spare_1_5 : Bool;
      Spare_1_6 : Bool;
      Spare_1_7 : Bool;
   END_STRUCT;

END_TYPE

TYPE "UDT_MCC_Status"
TITLE = UDT_Status_MCC
VERSION : 0.1
//Status of main control cabinet
//# Block Info
//- Title:            UDT_Status_MCC
//- Comment/Function: Status of main control cabinet
//- Library/Family:   APS
//- Author:           Jay Liu
//- Tested with:      ---
//- Engineering:      TIA Portal V20
//- Restrictions:     ---
//- Requirements:     ---
//
//# History
// |Version  | Date       | Author                 | Description                   |
// |---------|------------|------------------------|------------------------------ |
// |01.00.00 | 2026-01-22 | Jay Liu                | First released version        |
   STRUCT
      ER_Connection_Fault_AWCS : Bool;   // WCS communication error
      ER_Connection_Fault_SCADA : Bool;   // SCADA communication error
      ER_Connection_Fault_HMI : Bool;
      ER_Connection_Fault_Safety : Bool;
      ER_UR20_Not_Present : Bool;
      ER_UR20_Error : Bool;
      ER_UPS_Not_Present : Bool;
      ER_UPS_Error : Bool;
      ER_PAC3220_Not_Present : Bool;
      ER_PAC3220_Error : Bool;
      ER_XC216_Not_Present : Bool;
      ER_XC216_Error : Bool;
      WN_UPS_Battery_Low : Bool;
      WN_UPS_Battery_Change_Recommended : Bool;
      WN_UPS_Buffer_Mode_Active : Bool;
      WN_UPS_Battery_Connection_Down : Bool;
      WN_UPS_Input_Voltage_Fault : Bool;
      WN_UPS_Charge_Insufficient : Bool;
      WN_L1_N_Under_Voltage : Bool;
      WN_L1_N_Over_Voltage : Bool;
      WN_L2_N_Under_Voltage : Bool;
      WN_L2_N_Over_Voltage : Bool;
      WN_L3_N_Under_Voltage : Bool;
      WN_L3_N_Over_Voltage : Bool;
      WN_Unbalance_Voltage_Over_Limit : Bool;
      WN_Unbalance_Current_Over_Limit : Bool;
      WN_Cabinet_Temperature_High : Bool;
      ER_PowerSupply_NOK_G1011 : Bool;
      ER_PowerSupply_NOK_G1041 : Bool;
      ER_Main_Switch_Trip_Q1001 : Bool;
      ER_CB_F1011_Trip_Power_Supply : Bool;
      ER_CB_F1012_Trip_UPS_Out : Bool;
      ER_CB_F1021_Trip_HMI : Bool;
      ER_CB_F1022_Trip_CPU : Bool;
      ER_CB_F1023_Trip_XC216 : Bool;
      ER_CB_F1024_Trip_Safety_XC208 : Bool;
      ER_CB_F1025_Trip_Safety_CPU : Bool;
      ER_CB_F1026_Trip_Image_Server : Bool;
      ER_CB_F1031_Trip_Image_Switch : Bool;
      ER_CB_F1032_Trip_HLC_Gateway : Bool;
      ER_CB_F1033_Trip_Reserved : Bool;
      ER_CB_F1034_Trip_Reserved : Bool;
      ER_CB_F1072_Trip_PowerMeter_380VAC : Bool;
      ER_CB_F1072_Trip_PowerMeter_220VAC : Bool;
      ER_CB_F1041_Trip_Power_Supply : Bool;
      ER_CB_F105x_Trip_GC03_Scanner : Bool;
      ER_CB_F105x_Trip_GC04_Scanner : Bool;
      ER_CB_F105x_Trip_Safety_IO_24VDC : Bool;
      ER_CB_F105x_Trip_External_24VDC : Bool;
      ER_CB_F1081_Trip_AC01 : Bool;
      ER_CB_F1091_Trip_GC01_Inveter : Bool;
      ER_CB_F1092_Trip_AC02 : Bool;
      ER_CB_F1093_Trip_GC01_Interroll : Bool;
      ER_CB_F1094_Trip_GC01_SDC01 : Bool;
      ER_CB_F1101_Trip_GC02_Inveter : Bool;
      ER_CB_F1102_Trip_AC03 : Bool;
      ER_CB_F1103_Trip_Reversed : Bool;
      ER_CB_F1104_Trip_GC02_SDC01 : Bool;
      ER_CB_F1111_Trip_GC03_Inveter : Bool;
      ER_CB_F1112_Trip_AC04 : Bool;
      ER_CB_F1113_Trip_GC03_Interroll : Bool;
      ER_CB_F1114_Trip_GC03_SDC01 : Bool;
      ER_CB_F1115_Trip_GC03_SDC02 : Bool;
      ER_CB_F1121_Trip_GC04_Inveter : Bool;
      ER_CB_F1122_Trip_AC05 : Bool;
      ER_CB_F1123_Trip_Reversed : Bool;
      ER_CB_F1131_Trip_GC05_Inveter : Bool;
      ER_CB_F1132_Trip_GC05_Interroll : Bool;
      ER_CB_F1133_Trip_GC06_Inveter : Bool;
      ER_CB_F1134_Trip_GC06_Interroll : Bool;
      ER_CB_F1141_Trip_GC07_Inveter : Bool;
      ER_CB_F1142_Trip_GC07_Interroll : Bool;
      ER_CB_F1151_Trip_GC03_Inveter_Group2 : Bool;
      ER_CB_F1152_Trip_Reversed : Bool;
      ER_CB_F1153_Trip_Reversed : Bool;
      ER_CB_F1154_Trip_Reversed : Bool;
      ER_CB_F1155_Trip_EH01 : Bool;
      ER_CB_F1156_Trip_EH02 : Bool;
      ER_CB_F1157_Trip_EH03 : Bool;
      ER_CB_F1161_Trip_Fan : Bool;
      ER_CB_F1171_Trip_Socket : Bool;
      ER_KM_1641_Trip_GC01_Interroll : Bool;
      ER_KM_1642_Trip_GC01_Interroll : Bool;
      ER_KM_1643_Trip_Reversed : Bool;
      ER_KM_1644_Trip_Reversed : Bool;
      ER_KM_1645_Trip_GC03_Interroll : Bool;
      ER_KM_1646_Trip_GC03_Interroll : Bool;
      ER_KM_1647_Trip_Reversed : Bool;
      ER_KM_1648_Trip_Reversed : Bool;
      ER_KM_1651_Trip_GC05_Interroll : Bool;
      ER_KM_1652_Trip_GC05_Interroll : Bool;
      ER_KM_1653_Trip_GC05_Interroll : Bool;
      ER_KM_1654_Trip_GC05_Interroll : Bool;
      ER_KM_1655_Trip_GC05_Interroll : Bool;
      ER_KM_1656_Trip_GC05_Interroll : Bool;
      Spare_11_7 : Bool;
      Spare_12_0 : Bool;
      Spare_12_1 : Bool;
      Spare_12_2 : Bool;
      Spare_12_3 : Bool;
      Spare_12_4 : Bool;
      Spare_12_5 : Bool;
      Spare_12_6 : Bool;
      Spare_12_7 : Bool;
      Spare_13_0 : Bool;
      Spare_13_1 : Bool;
      Spare_13_2 : Bool;
      Spare_13_3 : Bool;
      Spare_13_4 : Bool;
      Spare_13_5 : Bool;
      Spare_13_6 : Bool;
      Spare_13_7 : Bool;
   END_STRUCT;

END_TYPE

TYPE "UDT_Echelon_Command"
VERSION : 0.1
   STRUCT
      Spare_0_0 : Bool;
      Spare_0_1 : Bool;
      Spare_0_2 : Bool;
      Spare_0_3 : Bool;
      Spare_0_4 : Bool;
      Spare_0_5 : Bool;
      Spare_0_6 : Bool;
      Spare_0_7 : Bool;
      Spare_1_0 : Bool;
      Spare_1_1 : Bool;
      Spare_1_2 : Bool;
      Spare_1_3 : Bool;
      Spare_1_4 : Bool;
      Spare_1_5 : Bool;
      Spare_1_6 : Bool;
      Spare_1_7 : Bool;
   END_STRUCT;

END_TYPE

TYPE "UDT_RLS_Interface"
VERSION : 0.1
   STRUCT
      Input : Struct
         Spare_0_0 : Bool;
         Spare_0_1 : Bool;
         Spare_0_2 : Bool;
         Spare_0_3 : Bool;
         Spare_0_4 : Bool;
         Spare_0_5 : Bool;
         Spare_0_6 : Bool;
         Spare_0_7 : Bool;
         Spare_1_0 : Bool;
         Spare_1_1 : Bool;
         Spare_1_2 : Bool;
         Spare_1_3 : Bool;
         Spare_1_4 : Bool;
         Spare_1_5 : Bool;
         Spare_1_6 : Bool;
         Spare_1_7 : Bool;
         Spare_Byte_2 : Byte;
         Spare_Byte_3 : Byte;
         Spare_Byte_4 : Byte;
         Spare_Byte_5 : Byte;
         Spare_Byte_6 : Byte;
         Spare_Byte_7 : Byte;
         Spare_Byte_8 : Byte;
         Spare_Byte_9 : Byte;
         Spare_Byte_10 : Byte;
         Spare_Byte_11 : Byte;
         Spare_Byte_12 : Byte;
         Spare_Byte_13 : Byte;
         Spare_Byte_14 : Byte;
         Spare_Byte_15 : Byte;
      END_STRUCT;
      Output : Struct
         Spare_0_0 : Bool;
         Spare_0_1 : Bool;
         Spare_0_2 : Bool;
         Spare_0_3 : Bool;
         Spare_0_4 : Bool;
         Spare_0_5 : Bool;
         Spare_0_6 : Bool;
         Spare_0_7 : Bool;
         Spare_1_0 : Bool;
         Spare_1_1 : Bool;
         Spare_1_2 : Bool;
         Spare_1_3 : Bool;
         Spare_1_4 : Bool;
         Spare_1_5 : Bool;
         Spare_1_6 : Bool;
         Spare_1_7 : Bool;
         Spare_Byte_2 : Byte;
         Spare_Byte_3 : Byte;
         Spare_Byte_4 : Byte;
         Spare_Byte_5 : Byte;
         Spare_Byte_6 : Byte;
         Spare_Byte_7 : Byte;
         Spare_Byte_8 : Byte;
         Spare_Byte_9 : Byte;
         Spare_Byte_10 : Byte;
         Spare_Byte_11 : Byte;
         Spare_Byte_12 : Byte;
         Spare_Byte_13 : Byte;
         Spare_Byte_14 : Byte;
         Spare_Byte_15 : Byte;
      END_STRUCT;
   END_STRUCT;

END_TYPE

TYPE "UDT_HMI_Command"
VERSION : 0.1
   STRUCT
      Start : Bool;
      Stop : Bool;
      Reset : Bool;
      Clear_Statistics : Bool;
   END_STRUCT;

END_TYPE

FUNCTION_BLOCK "FB_Conv_S210"
{ S7_Optimized_Access := 'TRUE' }
VERSION : 0.1
   VAR_INPUT
      i_Telegram_HW_ID { ExternalAccessible := 'False'; ExternalVisible := 'False'; ExternalWritable := 'False'} : HW_SUBMODULE;
      i_Additional_HW_ID { ExternalAccessible := 'False'; ExternalVisible := 'False'; ExternalWritable := 'False'} : HW_SUBMODULE;
      i_IO_PEC_Position : Bool;
      i_IO_PEC_Trigger : Bool;
      i_Setting : "UDT_Conv_S210_Setting";
      i_Command : "UDT_Conv_S210_Command";
      i_External_Request : "UDT_External_Request";
   END_VAR

   VAR_OUTPUT RETAIN
      o_Status : "UDT_Conv_S210_Status";
      o_General_Status : "UDT_General_Status";
      o_Diagnostics : "UDT_Conv_S210_Diagnostics";
   END_VAR

   VAR_IN_OUT
      io_Global : "UDT_Global";
      io_System_Control : "UDT_System_Control";
      io_S210_IO : "UDT_S210_HW_Interface";
      io_FIF_Upstream : "UDT_Flow_Interface";
      io_FIF : "UDT_Flow_Interface";
      io_FIF_Downstream : "UDT_Flow_Interface";
   END_VAR

   VAR
      s_FB_Displacement_AccDec : "FB_Displacement_AccDec";
      s_FB_EQP_PEC_Position : "FB_EQP_PEC_Position";
      s_FB_EQP_PEC_Trigger : "FB_EQP_PEC_Trigger";
      s_FB_EQP_Transport : "FB_EQP_Transport";
      s_FB_HW_Motor_S210 : "FB_HW_VFD_S210";
   END_VAR
   VAR RETAIN
      s_Cnt_PEC_Items { S7_SetPoint := 'True'} : Int;
      s_Speed_Select : Int;
      s_SW_Actual_Speed : Int;
      s_CMD_PEC_Preset_Latch : Bool;
      s_CMD_Motor : Bool;
      s_CMD_Motor_Reverse : Bool;
      s_HW_Req_Halt : Bool;
      s_PE_Position_Latch : Bool;
      s_PE_Trigger_Latch : Bool;
      s_Ext_Req_Stop : Bool;
      s_Ext_Req_Halt : Bool;
      s_Ext_Req_Disable_Send : Bool;
      s_Ext_Req_Disable_Recv : Bool;
      s_Ext_Req_Rest_ESave : Bool;
      s_Ext_Req_Clear_Data : Bool;
      s_SW_Motor_OnSpeed : Bool;
      s_HW_Motor_Running : Bool;
   END_VAR

   VAR_TEMP
      t_PEC_Position_Items : UDInt;
      t_PEC_Trigger_Items : UDInt;
      t_PEC_Position_Ready_To_Reset : Bool;
      t_PEC_Trigger_Ready_To_Reset : Bool;
      t_HW_VFD_Ready_To_Reset : Bool;
   END_VAR


BEGIN
	REGION NETWORK AA: Conveyor Cycle Displacement
	    IF NOT #i_Setting.Hardware.Use_Hardware_Feedback THEN
	        #s_FB_Displacement_AccDec(i_Conveyor_Speed   := #io_FIF.Speed,
	                                  i_Accelaration     := #i_Setting.Hardware.Acceleration,
	                                  i_Decelaration     := #i_Setting.Hardware.Deceleration,
	                                  i_Prev_Cycle_Time  := #io_Global.OB_Prev_Cycle_Time,
	                                  i_PPI_Displacement := 0,
	                                  i_Section_Run      := #io_FIF.Motor_Run,
	                                  o_Motor_On_Speed   => #o_General_Status.Motor_On_Speed,
	                                  o_Motor_Stopped    => #io_FIF.Motor_Stopped,
	                                  o_Actual_Speed     => #s_SW_Actual_Speed,
	                                  o_Displacement     => #io_FIF.Displacement);
	    ELSE
	        #o_General_Status.Motor_On_Speed := "FC_IsValue_InTolerance"(i_Value := #o_Diagnostics.Hardware.Actual_Speed,
	                                                                     i_Setpoint := #io_FIF.Speed,
	                                                                     i_High_Tolerance := -1,
	                                                                     i_Low_Tolerance := 10);
	        #io_FIF.Motor_Stopped := #o_Diagnostics.Hardware.Actual_Speed = 0;
	        #s_SW_Actual_Speed := #o_Diagnostics.Hardware.Actual_Speed;
	        #io_FIF.Displacement := #o_Diagnostics.Hardware.Actual_Displacement;
	    END_IF;

	    #o_General_Status.Motor_Stopped := #io_FIF.Motor_Stopped;
	END_REGION

	REGION NETWORK BA: Equipment layer - PEC
	    #s_FB_EQP_PEC_Position(i_IO_Available             := #io_System_Control.IO_Available,
	                           i_CMD_Reset                := #io_System_Control.OS_Reset_Jam,
	                           i_CMD_Clear_Stat           := #io_System_Control.OS_Clear_Statistics,
	                           i_CFG_Blockage_Length      := #i_Setting.PE1.Blockage_Length,
	                           i_CFG_Delay_On             := #i_Setting.PE1.Delay_On,
	                           i_CFG_Delay_Off            := #i_Setting.PE1.Delay_Off,
	                           i_CFG_Shifting_Offset      := #i_Setting.PE1.Shifting_Offset,
	                           i_CFG_Handover_Offset      := #i_Setting.PE1.Handover_Offset,
	                           i_CFG_Detect_PEC_OnStopped := #i_Setting.PE1.Detect_PEC_OnStopped,
	                           i_CFG_Reset_Block_PEC_Oc   := #i_Setting.PE1.Reset_Block_PEC_Oc,
	                           i_CFG_Item_On              := #i_Setting.PE1.Item_On,
	                           i_CMD_Preset_Latch         := #s_CMD_PEC_Preset_Latch,
	                           i_CMD_Clear_Data           := #s_Ext_Req_Clear_Data,
	                           i_Cycle_Count             := #io_FIF.Displacement,
	                           i_IO_PEC                   := #i_IO_PEC_Position,
	                           i_Section_Running          := NOT #io_FIF.Motor_Stopped,
	                           o_Ready_To_Reset           => #t_PEC_Position_Ready_To_Reset,
	                           o_ER_PEC_Blockage          => #o_Status.ER_PE1_Blockage,
	                           o_PEC_Filter               => #s_PE_Position_Latch,
	                           o_Handover                 => #io_FIF.Handover,
	                           o_Cnt_Buffer_Used          => #s_Cnt_PEC_Items,
	                           o_Stat_Items               => #t_PEC_Position_Items);

	    #s_FB_EQP_PEC_Trigger(i_IO_Available             := #io_System_Control.IO_Available,
	                          i_CMD_Reset                := #io_System_Control.OS_Reset_Jam,
	                          i_CMD_Clear_Stat           := #io_System_Control.OS_Clear_Statistics,
	                          i_CFG_Blockage_Length      := #i_Setting.PE2.Blockage_Length,
	                          i_CFG_Delay_On             := #i_Setting.PE2.Delay_On,
	                          i_CFG_Delay_Off            := #i_Setting.PE2.Delay_Off,
	                          i_CFG_Detect_PEC_OnStopped := #i_Setting.PE2.Detect_PEC_OnStopped,
	                          i_CFG_Reset_Block_PEC_Oc   := #i_Setting.PE2.Reset_Block_PEC_Oc,
	                          i_CFG_Item_On              := #i_Setting.PE2.Item_On,
	                          i_CMD_Preset_Latch         := FALSE,
	                          i_Cycle_Count             := #io_FIF.Displacement,
	                          i_IO_PEC                   := #i_IO_PEC_Trigger,
	                          i_Section_Running          := NOT #io_FIF.Motor_Stopped,
	                          o_Ready_To_Reset           => #t_PEC_Trigger_Ready_To_Reset,
	                          o_ER_PEC_Blockage          => #o_Status.ER_PE2_Blockage,
	                          o_PEC_Filter               => #s_PE_Trigger_Latch,
	                          o_Stat_Items               => #t_PEC_Trigger_Items);

	    #io_FIF.PECTrigger_Latch := #s_PE_Trigger_Latch;
	END_REGION

	REGION NETWORK CA: Conditions to basic control
	    // Condition to request stop
	    #s_Ext_Req_Stop := #o_Status.ER_Servo_PN_NotPresent
	    //OR #o_Status.ER_Motor_PN_Error
	    OR #o_Status.ER_Servo_Fault
	    OR #o_Status.ER_Servo_STO_Active
	    OR #i_External_Request.Request_Stop;

	    // Condition to request halt
	    #s_Ext_Req_Halt := #s_HW_Req_Halt OR #i_External_Request.Request_Halt OR #i_Command.Man_Mode OR #o_Status.ER_PE1_Blockage OR #o_Status.ER_PE2_Blockage;

	    // Condition to request disable send
	    #s_Ext_Req_Disable_Send := #i_External_Request.Request_Disable_Send;

	    // Condition to request disable receive
	    #s_Ext_Req_Disable_Recv := #i_External_Request.Request_Disable_Receive OR #i_Command.Man_Mode;

	    // Condition to request reset engergy saving
	    #s_Ext_Req_Rest_ESave := #i_External_Request.Request_Reset_EnergySave OR #io_Global.Common_Setting.Disable_Energy_Saving OR #i_Command.Cmd_Reset_ESave;

	    // Condition to request clear flow interface data
	    #s_Ext_Req_Clear_Data := #i_External_Request.Request_Clear_Data OR (#i_Command.Man_Clear AND #i_Command.Man_Mode);
	END_REGION

	REGION NETWORK DA: Equipment Layer - Basic
	    #s_FB_EQP_Transport(i_Enable                 := #io_System_Control.Enable,
	                        i_IO_Available           := #io_System_Control.IO_Available,
	                        i_Safety_OK              := #io_System_Control.Safety_OK,
	                        i_CMD_Reset              := #io_System_Control.OS_Reset,
	                        i_CMD_Start              := #io_System_Control.OS_Start,
	                        i_CMD_Controlled_Stop    := #io_System_Control.Controlled_Stop,
	                        i_End_PEC_Latch          := #s_PE_Position_Latch,
	                        i_Manual_Run             := #i_Command.Man_Run AND #i_Command.Man_Mode,
	                        i_CFG_Slave_Conveyor     := #i_Setting.Base_Conveyor.Slave_Mode,
	                        i_CFG_Enable_DieForward  := #i_Setting.Base_Conveyor.Enable_DieForward,
	                        i_Delay_Waiting_Item     := #i_Setting.Base_Conveyor.Delay_Waiting_Item,
	                        i_Delay_Dieback          := #i_Setting.Base_Conveyor.Delay_Dieback,
	                        i_Delay_Startup          := #i_Setting.Base_Conveyor.Delay_Startup,
	                        i_Delay_Finish_Handover  := #i_Setting.Base_Conveyor.Delay_Finish_Handover,
	                        i_Delay_Energysave       := #i_Setting.Base_Conveyor.Delay_Energysave,
	                        i_Delay_Cascade_Startup  := #i_Setting.Base_Conveyor.Delay_Cascade_Startup,
	                        i_Delay_Cascade_Shutdown := #i_Setting.Base_Conveyor.Delay_Cascade_Shutdown,
	                        i_Delay_Motor_Startup    := 0,
	                        i_Minimum_Gap            := #i_Setting.Flow_Control.Minimum_Gap,
	                        i_Minimum_Head_To_Head   := #i_Setting.Flow_Control.Minimum_Head_To_Head,
	                        i_Ext_Req_Stop           := #s_Ext_Req_Stop,
	                        i_Ext_Req_Halt           := #s_Ext_Req_Halt,
	                        i_Ext_Req_Dis_Send       := #s_Ext_Req_Disable_Send,
	                        i_Ext_Req_Dis_Recv       := #s_Ext_Req_Disable_Recv,
	                        i_Ext_Req_Rst_ESave      := #s_Ext_Req_Rest_ESave,
	                        i_Ext_Req_Clear_Data     := #s_Ext_Req_Clear_Data,
	                        o_Ready_To_Start         => #io_System_Control.Ready_To_Start,
	                        o_ST_Safety_Stop         => #o_General_Status.Safety_Stop,
	                        o_ST_Items               => #o_General_Status.Items,
	                        o_ST_Die_Back            => #o_General_Status.Die_Back,
	                        o_ST_Motor_Running       => #o_General_Status.Motor_Running,
	                        o_ST_Started             => #o_General_Status.Started,
	                        o_ST_Energy_Saving       => #o_General_Status.Energy_Saving,
	                        o_MTR_Run                => #s_CMD_Motor,
	                        io_Global                := #io_Global,
	                        io_FIF_Upstream          := #io_FIF_Upstream,
	                        io_FIF                   := #io_FIF,
	                        io_FIF_Downstream        := #io_FIF_Downstream);
	END_REGION

	REGION NETWORK EA: Hardware Layer - S210 Servo
	    #s_Speed_Select := #i_External_Request.Request_Speed;

	    #s_FB_HW_Motor_S210(i_Telegram_HW_ID        := #i_Telegram_HW_ID,
	                        i_Additional_HW_ID      := #i_Additional_HW_ID,
	                        i_Enable                := (#io_System_Control.Enable OR #i_Command.Man_Mode) AND NOT #i_Command.Man_DisableAxis,
	                        i_IO_Available          := #io_System_Control.IO_Available,
	                        i_Safety_OK             := #io_System_Control.Safety_OK,
	                        i_CMD_Reset             := #io_System_Control.OS_Reset,
	                        i_CMD_Clear_Stat        := #io_System_Control.OS_Clear_Statistics,
	                        i_HW_Setting            := #i_Setting.Hardware,
	                        i_CFG_Motor_Switch_Time := 200,
	                        i_CMD_Select_Speed      := #s_Speed_Select,
	                        i_CMD_Motor_Run         := #s_CMD_Motor,
	                        i_CMD_Motor_Reverse     := #s_CMD_Motor_Reverse,
	                        o_Ready_To_Reset        => #t_HW_VFD_Ready_To_Reset,
	                        o_Req_Halt              => #s_HW_Req_Halt,
	                        o_ER_PN_Not_Present     => #o_Status.ER_Servo_PN_NotPresent,
	                        o_ER_PN_Error           => #o_Status.ER_Servo_PN_Error,
	                        o_ER_Motor_Fault        => #o_Status.ER_Servo_Fault,
	                        o_WN_Motor_Alarm        => #o_Status.WN_Servo_Alarm,
	                        o_ER_STO_Active         => #o_Status.ER_Servo_STO_Active,
	                        o_ST_Motor_Running      => #s_HW_Motor_Running,
	                        o_FaultCode             => #o_Status.FaultCode,
	                        o_AlarmCode             => #o_Status.AlarmCode,
	                        o_Speed_Selected        => #io_FIF.Speed,
	                        o_Diagnostics           => #o_Diagnostics.Hardware,
	                        io_Global               := #io_Global,
	                        io_S210_Interface       := #io_S210_IO);
	END_REGION

	REGION NETWORK: Diagnositcs
	    #o_Diagnostics.RTS := #io_FIF.RTS;
	    #o_Diagnostics.TIP := #io_FIF.TIP;
	    #o_Diagnostics.Downstream_RTR := #io_FIF_Downstream.RTR;
	    #o_Diagnostics.Displacement := #io_FIF.Displacement;
	    #o_Diagnostics.Items_Count := MAX_UDINT(IN1 := #t_PEC_Position_Items, IN2 := #t_PEC_Trigger_Items);
	END_REGION

	REGION NETWORK FA: Make Generate Status
	    #o_Status.OL_Maintenance_Mode := #i_Command.Man_Mode;

	    #o_General_Status.Safety_Stop := #o_Status.ER_Servo_STO_Active OR NOT #io_System_Control.Safety_OK;
	    #o_General_Status.Off_Line := #o_Status.OL_Maintenance_Mode;
	    #o_General_Status.Manual := FALSE;
	    #o_General_Status.Error := #o_Status.ER_Servo_PN_NotPresent
	    //OR #o_Status.ER_Motor_PN_Error
	    OR #o_Status.ER_Servo_Fault;
	    #o_General_Status.Jam := #o_Status.ER_PE1_Blockage OR #o_Status.ER_PE2_Blockage;
	    #o_General_Status.Warning := #o_Status.WN_Servo_Alarm;

	END_REGION

	REGION NETWORK EA: System Feedback State
	    #io_System_Control.Ready_To_Reset := #t_PEC_Position_Ready_To_Reset
	    OR #t_PEC_Trigger_Ready_To_Reset
	    OR #t_HW_VFD_Ready_To_Reset;
	END_REGION
END_FUNCTION_BLOCK

FUNCTION_BLOCK "FB_Conv_G115D"
{ S7_Optimized_Access := 'TRUE' }
VERSION : 0.1
   VAR_INPUT
      i_Telegram_HW_ID : HW_SUBMODULE;
      i_Additional_HW_ID : HW_SUBMODULE;
      i_IO_PEC_Position : Bool;
      i_IO_PEC_Trigger : Bool;
      i_Setting : "UDT_Conv_G115D_Setting";
      i_External_Request : "UDT_External_Request";
      i_Command : "UDT_Conv_G115D_Command";
   END_VAR

   VAR_OUTPUT RETAIN
      o_Status : "UDT_Conv_G115D_Status";
      o_General_Status : "UDT_General_Status";
      o_Diagnostics : "UDT_Conv_G115D_Diagnostics";
   END_VAR

   VAR_IN_OUT
      io_Global : "UDT_Global";
      io_System_Control : "UDT_System_Control";
      io_G115D_IO : "UDT_G115D_HW_Interface";
      io_FIF_Upstream : "UDT_Flow_Interface";
      io_FIF : "UDT_Flow_Interface";
      io_FIF_Downstream : "UDT_Flow_Interface";
   END_VAR

   VAR
      s_FB_Displacement_AccDec : "FB_Displacement_AccDec";
      s_FB_EQP_PEC_Position : "FB_EQP_PEC_Position";
      s_FB_EQP_PEC_Trigger : "FB_EQP_PEC_Trigger";
      s_FB_EQP_Transport : "FB_EQP_Transport";
      s_FB_HW_VFD_G115D : "FB_HW_VFD_G115D";
   END_VAR
   VAR RETAIN
      s_Cnt_PEC_Items : Int;
      s_Speed_Select : Int;
      s_SW_Actual_Speed : Int;
      s_HW_Actual_Speed : Int;
      s_CMD_PEC_Preset_Latch : Bool;
      s_CMD_Motor : Bool;
      s_CMD_Motor_Reverse : Bool;
      s_HW_Req_Halt : Bool;
      s_PE_Position_Latch : Bool;
      s_PE_Trigger_Latch : Bool;
      s_Ext_Req_Stop : Bool;
      s_Ext_Req_Halt : Bool;
      s_Ext_Req_Disable_Send : Bool;
      s_Ext_Req_Disable_Recv : Bool;
      s_Ext_Req_Rest_ESave : Bool;
      s_Ext_Req_Clear_Data : Bool;
      s_SW_Motor_OnSpeed : Bool;
      s_HW_Motor_Running : Bool;
   END_VAR

   VAR_TEMP
      t_PEC_Position_Items : UDInt;
      t_PEC_Trigger_Items : UDInt;
      t_PEC_Position_Ready_To_Reset : Bool;
      t_PEC_Trigger_Ready_To_Reset : Bool;
      t_HW_VFD_Ready_To_Reset : Bool;
   END_VAR


BEGIN
	REGION NETWORK AA: Conveyor Cycle Displacement
	    #s_FB_Displacement_AccDec(i_Conveyor_Speed   := #io_FIF.Speed,
	                              i_Accelaration     := #i_Setting.Hardware.Acceleration,
	                              i_Decelaration     := #i_Setting.Hardware.Deceleration,
	                              i_Prev_Cycle_Time  := #io_Global.OB_Prev_Cycle_Time,
	                              i_PPI_Displacement := 0,
	                              i_Section_Run      := #io_FIF.Motor_Run,
	                              o_Motor_On_Speed   => #o_General_Status.Motor_On_Speed,
	                              o_Motor_Stopped    => #io_FIF.Motor_Stopped,
	                              o_Actual_Speed     => #s_SW_Actual_Speed,
	                              o_Displacement     => #io_FIF.Displacement);

	    #o_General_Status.Motor_Stopped := #io_FIF.Motor_Stopped;
	END_REGION

	REGION NETWORK BA: Equipment layer - PEC
	    #s_FB_EQP_PEC_Position(i_IO_Available             := #io_System_Control.IO_Available,
	                           i_CMD_Reset                := #io_System_Control.OS_Reset_Jam,
	                           i_CMD_Clear_Stat           := #io_System_Control.OS_Clear_Statistics,
	                           i_CFG_Blockage_Length      := #i_Setting.PE1.Blockage_Length,
	                           i_CFG_Delay_On             := #i_Setting.PE1.Delay_On,
	                           i_CFG_Delay_Off            := #i_Setting.PE1.Delay_Off,
	                           i_CFG_Shifting_Offset      := #i_Setting.PE1.Shifting_Offset,
	                           i_CFG_Handover_Offset      := #i_Setting.PE1.Handover_Offset,
	                           i_CFG_Detect_PEC_OnStopped := #i_Setting.PE1.Detect_PEC_OnStopped,
	                           i_CFG_Reset_Block_PEC_Oc   := #i_Setting.PE1.Reset_Block_PEC_Oc,
	                           i_CFG_Item_On              := #i_Setting.PE1.Item_On,
	                           i_CMD_Preset_Latch         := #s_CMD_PEC_Preset_Latch,
	                           i_CMD_Clear_Data           := #s_Ext_Req_Clear_Data,
	                           i_Cycle_Count              := #io_FIF.Displacement,
	                           i_IO_PEC                   := #i_IO_PEC_Position,
	                           i_Section_Running          := NOT #io_FIF.Motor_Stopped,
	                           o_Ready_To_Reset           => #t_PEC_Position_Ready_To_Reset,
	                           o_ER_PEC_Blockage          => #o_Status.ER_PE1_Blockage,
	                           o_PEC_Filter               => #s_PE_Position_Latch,
	                           o_Handover                 => #io_FIF.Handover,
	                           o_Cnt_Buffer_Used          => #s_Cnt_PEC_Items,
	                           o_Stat_Items               => #t_PEC_Position_Items);

	    #s_FB_EQP_PEC_Trigger(i_IO_Available             := #io_System_Control.IO_Available,
	                          i_CMD_Reset                := #io_System_Control.OS_Reset_Jam,
	                          i_CMD_Clear_Stat           := #io_System_Control.OS_Clear_Statistics,
	                          i_CFG_Blockage_Length      := #i_Setting.PE2.Blockage_Length,
	                          i_CFG_Delay_On             := #i_Setting.PE2.Delay_On,
	                          i_CFG_Delay_Off            := #i_Setting.PE2.Delay_Off,
	                          i_CFG_Detect_PEC_OnStopped := #i_Setting.PE2.Detect_PEC_OnStopped,
	                          i_CFG_Reset_Block_PEC_Oc   := #i_Setting.PE2.Reset_Block_PEC_Oc,
	                          i_CFG_Item_On              := #i_Setting.PE2.Item_On,
	                          i_CMD_Preset_Latch         := false,
	                          i_Cycle_Count              := #io_FIF.Displacement,
	                          i_IO_PEC                   := #i_IO_PEC_Trigger,
	                          i_Section_Running          := NOT #io_FIF.Motor_Stopped,
	                          o_Ready_To_Reset           => #t_PEC_Trigger_Ready_To_Reset,
	                          o_ER_PEC_Blockage          => #o_Status.ER_PE2_Blockage,
	                          o_PEC_Filter               => #s_PE_Trigger_Latch,
	                          o_Stat_Items               => #t_PEC_Trigger_Items);

	    #io_FIF.PECTrigger_Latch := #s_PE_Trigger_Latch;
	END_REGION

	REGION NETWORK CA: Conditions to basic control
	    // Condition to request stop
	    #s_Ext_Req_Stop := #o_Status.ER_VFD_PN_NotPresent
	    //OR #o_Status.ER_Motor_PN_Error
	    OR #o_Status.ER_VFD_Fault
	    OR #o_Status.ER_VFD_STO_Active
	    OR #i_External_Request.Request_Stop;

	    // Condition to request halt
	    #s_Ext_Req_Halt := #s_HW_Req_Halt OR #i_External_Request.Request_Halt OR #i_Command.Man_Mode OR #o_Status.ER_PE1_Blockage OR #o_Status.ER_PE2_Blockage;

	    // Condition to request disable send
	    #s_Ext_Req_Disable_Send := #i_External_Request.Request_Disable_Send;

	    // Condition to request disable receive
	    #s_Ext_Req_Disable_Recv := #i_External_Request.Request_Disable_Receive OR #i_Command.Man_Mode;

	    // Condition to request reset engergy saving
	    #s_Ext_Req_Rest_ESave := #i_External_Request.Request_Reset_EnergySave OR #io_Global.Common_Setting.Disable_Energy_Saving OR #i_Command.Cmd_Reset_ESave OR #s_PE_Trigger_Latch OR #s_FB_EQP_PEC_Position.s_PEC_Filter;

	    // Condition to request clear flow interface data
	    #s_Ext_Req_Clear_Data := #i_External_Request.Request_Clear_Data OR (#i_Command.Man_Clear AND #i_Command.Man_Mode);
	END_REGION

	REGION NETWORK DA: Equipment Layer - Basic
	    #s_FB_EQP_Transport(i_Enable                 := #io_System_Control.Enable,
	                        i_IO_Available           := #io_System_Control.IO_Available,
	                        i_Safety_OK              := #io_System_Control.Safety_OK,
	                        i_CMD_Reset              := #io_System_Control.OS_Reset,
	                        i_CMD_Start              := #io_System_Control.OS_Start,
	                        i_CMD_Controlled_Stop    := #io_System_Control.Controlled_Stop,
	                        i_End_PEC_Latch          := #s_PE_Position_Latch,
	                        i_Manual_Run             := #i_Command.Man_Run AND #i_Command.Man_Mode,
	                        i_CFG_Slave_Conveyor     := #i_Setting.Base_Conveyor.Slave_Mode,
	                        i_CFG_Enable_DieForward  := #i_Setting.Base_Conveyor.Enable_DieForward,
	                        i_Delay_Waiting_Item     := #i_Setting.Base_Conveyor.Delay_Waiting_Item,
	                        i_Delay_Dieback          := #i_Setting.Base_Conveyor.Delay_Dieback,
	                        i_Delay_Startup          := #i_Setting.Base_Conveyor.Delay_Startup,
	                        i_Delay_Finish_Handover  := #i_Setting.Base_Conveyor.Delay_Finish_Handover,
	                        i_Delay_Energysave       := #i_Setting.Base_Conveyor.Delay_Energysave,
	                        i_Delay_Cascade_Startup  := #i_Setting.Base_Conveyor.Delay_Cascade_Startup,
	                        i_Delay_Cascade_Shutdown := #i_Setting.Base_Conveyor.Delay_Cascade_Shutdown,
	                        i_Delay_Motor_Startup    := #i_Setting.Hardware.Magnetization_Delay,
	                        i_Minimum_Gap            := #i_Setting.Flow_Control.Minimum_Gap,
	                        i_Minimum_Head_To_Head   := #i_Setting.Flow_Control.Minimum_Head_To_Head,
	                        i_Ext_Req_Stop           := #s_Ext_Req_Stop,
	                        i_Ext_Req_Halt           := #s_Ext_Req_Halt,
	                        i_Ext_Req_Dis_Send       := #s_Ext_Req_Disable_Send,
	                        i_Ext_Req_Dis_Recv       := #s_Ext_Req_Disable_Recv,
	                        i_Ext_Req_Rst_ESave      := #s_Ext_Req_Rest_ESave,
	                        i_Ext_Req_Clear_Data     := #s_Ext_Req_Clear_Data,
	                        o_Ready_To_Start         => #io_System_Control.Ready_To_Start,
	                        o_ST_Safety_Stop         => #o_General_Status.Safety_Stop,
	                        o_ST_Items               => #o_General_Status.Items,
	                        o_ST_Die_Back            => #o_General_Status.Die_Back,
	                        o_ST_Motor_Running       => #o_General_Status.Motor_Running,
	                        o_ST_Started             => #o_General_Status.Started,
	                        o_ST_Energy_Saving       => #o_General_Status.Energy_Saving,
	                        o_MTR_Run                => #s_CMD_Motor,
	                        io_Global                := #io_Global,
	                        io_FIF_Upstream          := #io_FIF_Upstream,
	                        io_FIF                   := #io_FIF,
	                        io_FIF_Downstream        := #io_FIF_Downstream);
	END_REGION

	REGION NETWORK EA: Hardware Layer - G115D Convertor
	    #s_Speed_Select := #i_External_Request.Request_Speed;

	    #s_FB_HW_VFD_G115D(i_Telegram_HW_ID        := #i_Telegram_HW_ID,
	                       i_Additional_HW_ID      := #i_Additional_HW_ID,
	                       i_Enable                := (#io_System_Control.Enable OR #i_Command.Man_Mode) AND NOT #i_Command.Man_DisableAxis,
	                       i_IO_Available          := #io_System_Control.IO_Available,
	                       i_Safety_OK             := #io_System_Control.Safety_OK,
	                       i_CMD_Reset             := #io_System_Control.OS_Reset,
	                       i_CMD_Clear_Stat        := #io_System_Control.OS_Clear_Statistics,
	                       i_HW_Setting            := #i_Setting.Hardware,
	                       i_CFG_Motor_Switch_Time := 500,
	                       i_CMD_Select_Speed      := #s_Speed_Select,
	                       i_CMD_Motor_Run         := #s_CMD_Motor,
	                       i_CMD_Motor_Reverse     := #s_CMD_Motor_Reverse,
	                       o_Ready_To_Reset        => #t_HW_VFD_Ready_To_Reset,
	                       o_Req_Halt              => #s_HW_Req_Halt,
	                       o_ER_PN_Not_Present     => #o_Status.ER_VFD_PN_NotPresent,
	                       o_ER_PN_Error           => #o_Status.ER_VFD_PN_Error,
	                       o_ER_Motor_Fault        => #o_Status.ER_VFD_Fault,
	                       o_WN_Motor_Alarm        => #o_Status.WN_VFD_Alarm,
	                       o_ER_STO_Active         => #o_Status.ER_VFD_STO_Active,
	                       o_WN_No_MemoryCard      => #o_Status.WN_No_MemoryCard,
	                       o_ST_Motor_Running      => #s_HW_Motor_Running,
	                       o_FaultCode             => #o_Status.FaultCode,
	                       o_AlarmCode             => #o_Status.AlarmCode,
	                       o_Speed_Selected        => #io_FIF.Speed,
	                       o_Diagnostics           => #o_Diagnostics.Hardware,
	                       io_Global               := #io_Global,
	                       io_G115D_Interface      := #io_G115D_IO);
	END_REGION

	REGION NETWORK: Diagnositcs
	    #o_Diagnostics.RTS := #io_FIF.RTS;
	    #o_Diagnostics.TIP := #io_FIF.TIP;
	    #o_Diagnostics.Downstream_RTR := #io_FIF_Downstream.RTR;
	    #o_Diagnostics.Displacement := #io_FIF.Displacement;
	    #o_Diagnostics.Items_Count := MAX_UDINT(IN1 := #t_PEC_Position_Items, IN2 := #t_PEC_Trigger_Items);
	END_REGION

	REGION NETWORK FA: Make Generate Status
	    #o_Status.OL_Maintenance_Mode := #i_Command.Man_Mode;

	    #o_General_Status.Safety_Stop := #o_Status.ER_VFD_STO_Active OR NOT #io_System_Control.Safety_OK;
	    #o_General_Status.Off_Line := #o_Status.OL_Maintenance_Mode;
	    #o_General_Status.Manual := FALSE;
	    #o_General_Status.Error := #o_Status.ER_VFD_PN_NotPresent
	    OR #o_Status.ER_VFD_PN_Error
	    OR #o_Status.ER_VFD_Fault;
	    #o_General_Status.Jam := #o_Status.ER_PE1_Blockage OR #o_Status.ER_PE2_Blockage;
	    #o_General_Status.Warning := #o_Status.WN_VFD_Alarm OR #o_Status.WN_No_MemoryCard;
	END_REGION

	REGION NETWORK EA: System Feedback State
	    #io_System_Control.Ready_To_Reset := #t_PEC_Position_Ready_To_Reset
	    OR #t_PEC_Trigger_Ready_To_Reset
	    OR #t_HW_VFD_Ready_To_Reset;
	END_REGION
END_FUNCTION_BLOCK

TYPE "UDT_PAC_HW_Interface"
VERSION : 0.1
   STRUCT
      Input { S7_SetPoint := 'False'} : "UDT_PAC_HW_Input";
      Output : "UDT_PAC_HW_Output";
   END_STRUCT;

END_TYPE

TYPE "UDT_AC01_IO"
VERSION : 0.1
   STRUCT
      Input : Struct
         Spare_0_0 : Bool;
         Spare_0_1 : Bool;
         Spare_0_2 : Bool;
         Spare_0_3 : Bool;
         Spare_0_4 : Bool;
         Spare_0_5 : Bool;
         Spare_0_6 : Bool;
         Spare_0_7 : Bool;
         Spare_1_0 : Bool;
         Spare_1_1 : Bool;
         Spare_1_2 : Bool;
         Spare_1_3 : Bool;
         Spare_1_4 : Bool;
         Spare_1_5 : Bool;
         Spare_1_6 : Bool;
         Spare_1_7 : Bool;
      END_STRUCT;
      Output : Struct
         Spare_0_0 : Bool;
         Spare_0_1 : Bool;
         Spare_0_2 : Bool;
         Spare_0_3 : Bool;
         Spare_0_4 : Bool;
         Spare_0_5 : Bool;
         Spare_0_6 : Bool;
         Spare_0_7 : Bool;
         Spare_1_0 : Bool;
         Spare_1_1 : Bool;
         Spare_1_2 : Bool;
         Spare_1_3 : Bool;
         Spare_1_4 : Bool;
         Spare_1_5 : Bool;
         Spare_1_6 : Bool;
         Spare_1_7 : Bool;
      END_STRUCT;
   END_STRUCT;

END_TYPE

TYPE "UDT_AC02_IO"
VERSION : 0.1
   STRUCT
      Input : Struct
         Spare_0_0 : Bool;
         Spare_0_1 : Bool;
         Spare_0_2 : Bool;
         Spare_0_3 : Bool;
         Spare_0_4 : Bool;
         Spare_0_5 : Bool;
         Spare_0_6 : Bool;
         Spare_0_7 : Bool;
         Spare_1_0 : Bool;
         Spare_1_1 : Bool;
         Spare_1_2 : Bool;
         Spare_1_3 : Bool;
         Spare_1_4 : Bool;
         Spare_1_5 : Bool;
         Spare_1_6 : Bool;
         Spare_1_7 : Bool;
      END_STRUCT;
      Output : Struct
         Spare_0_0 : Bool;
         Spare_0_1 : Bool;
         Spare_0_2 : Bool;
         Spare_0_3 : Bool;
         Spare_0_4 : Bool;
         Spare_0_5 : Bool;
         Spare_0_6 : Bool;
         Spare_0_7 : Bool;
         Spare_1_0 : Bool;
         Spare_1_1 : Bool;
         Spare_1_2 : Bool;
         Spare_1_3 : Bool;
         Spare_1_4 : Bool;
         Spare_1_5 : Bool;
         Spare_1_6 : Bool;
         Spare_1_7 : Bool;
      END_STRUCT;
   END_STRUCT;

END_TYPE

TYPE "UDT_AC03_IO"
VERSION : 0.1
   STRUCT
      Input : Struct
         Spare_0_0 : Bool;
         Spare_0_1 : Bool;
         Spare_0_2 : Bool;
         Spare_0_3 : Bool;
         Spare_0_4 : Bool;
         Spare_0_5 : Bool;
         Spare_0_6 : Bool;
         Spare_0_7 : Bool;
         Spare_1_0 : Bool;
         Spare_1_1 : Bool;
         Spare_1_2 : Bool;
         Spare_1_3 : Bool;
         Spare_1_4 : Bool;
         Spare_1_5 : Bool;
         Spare_1_6 : Bool;
         Spare_1_7 : Bool;
      END_STRUCT;
      Output : Struct
         Spare_0_0 : Bool;
         Spare_0_1 : Bool;
         Spare_0_2 : Bool;
         Spare_0_3 : Bool;
         Spare_0_4 : Bool;
         Spare_0_5 : Bool;
         Spare_0_6 : Bool;
         Spare_0_7 : Bool;
         Spare_1_0 : Bool;
         Spare_1_1 : Bool;
         Spare_1_2 : Bool;
         Spare_1_3 : Bool;
         Spare_1_4 : Bool;
         Spare_1_5 : Bool;
         Spare_1_6 : Bool;
         Spare_1_7 : Bool;
      END_STRUCT;
   END_STRUCT;

END_TYPE

TYPE "UDT_AC04_IO"
VERSION : 0.1
   STRUCT
      Input : Struct
         Spare_0_0 : Bool;
         Spare_0_1 : Bool;
         Spare_0_2 : Bool;
         Spare_0_3 : Bool;
         Spare_0_4 : Bool;
         Spare_0_5 : Bool;
         Spare_0_6 : Bool;
         Spare_0_7 : Bool;
         Spare_1_0 : Bool;
         Spare_1_1 : Bool;
         Spare_1_2 : Bool;
         Spare_1_3 : Bool;
         Spare_1_4 : Bool;
         Spare_1_5 : Bool;
         Spare_1_6 : Bool;
         Spare_1_7 : Bool;
      END_STRUCT;
      Output : Struct
         Spare_0_0 : Bool;
         Spare_0_1 : Bool;
         Spare_0_2 : Bool;
         Spare_0_3 : Bool;
         Spare_0_4 : Bool;
         Spare_0_5 : Bool;
         Spare_0_6 : Bool;
         Spare_0_7 : Bool;
         Spare_1_0 : Bool;
         Spare_1_1 : Bool;
         Spare_1_2 : Bool;
         Spare_1_3 : Bool;
         Spare_1_4 : Bool;
         Spare_1_5 : Bool;
         Spare_1_6 : Bool;
         Spare_1_7 : Bool;
      END_STRUCT;
   END_STRUCT;

END_TYPE

TYPE "UDT_AC05_IO"
VERSION : 0.1
   STRUCT
      Input : Struct
         Spare_0_0 : Bool;
         Spare_0_1 : Bool;
         Spare_0_2 : Bool;
         Spare_0_3 : Bool;
         Spare_0_4 : Bool;
         Spare_0_5 : Bool;
         Spare_0_6 : Bool;
         Spare_0_7 : Bool;
         Spare_1_0 : Bool;
         Spare_1_1 : Bool;
         Spare_1_2 : Bool;
         Spare_1_3 : Bool;
         Spare_1_4 : Bool;
         Spare_1_5 : Bool;
         Spare_1_6 : Bool;
         Spare_1_7 : Bool;
      END_STRUCT;
      Output : Struct
         Spare_0_0 : Bool;
         Spare_0_1 : Bool;
         Spare_0_2 : Bool;
         Spare_0_3 : Bool;
         Spare_0_4 : Bool;
         Spare_0_5 : Bool;
         Spare_0_6 : Bool;
         Spare_0_7 : Bool;
         Spare_1_0 : Bool;
         Spare_1_1 : Bool;
         Spare_1_2 : Bool;
         Spare_1_3 : Bool;
         Spare_1_4 : Bool;
         Spare_1_5 : Bool;
         Spare_1_6 : Bool;
         Spare_1_7 : Bool;
      END_STRUCT;
   END_STRUCT;

END_TYPE

TYPE "UDT_SDC_4Servos_IO"
VERSION : 0.1
   STRUCT
      Spare_0_0 : Bool;
      Spare_0_1 : Bool;
      Spare_0_2 : Bool;
      Spare_0_3 : Bool;
      Spare_0_4 : Bool;
      Spare_0_5 : Bool;
      Spare_0_6 : Bool;
      Spare_0_7 : Bool;
      Spare_1_0 : Bool;
      Spare_1_1 : Bool;
      Spare_1_2 : Bool;
      Spare_1_3 : Bool;
      Spare_1_4 : Bool;
      Spare_1_5 : Bool;
      Spare_1_6 : Bool;
      Spare_1_7 : Bool;
   END_STRUCT;

END_TYPE

TYPE "UDT_Conv_Multiple_S210_Status"
VERSION : 0.1
   STRUCT
      OL_Maintenance_Mode : Bool;   // Maintenance mode on
      ER_PE1_Blockage : Bool;   // PE1 blockage
      ER_PE2_Blockage : Bool;   // PE2 blockage
      ER_U01_Servo_PN_NotPresent : Bool;   // Servo driver not present on profinet network
      ER_U01_Servo_PN_Error : Bool;   // Servo driver has error profinet network
      ER_U01_Servo_Fault : Bool;   // Servo driver has error
      WN_U01_Servo_Alarm : Bool;   // Servo driver has an warning
      ER_U01_Servo_STO_Active : Bool;   // Servo driver STO is active
      WN_U01_No_MemoryCard : Bool;   // Memory card is missing
      ER_U02_Servo_PN_NotPresent : Bool;   // Servo driver not present on profinet network
      ER_U02_Servo_PN_Error : Bool;   // Servo driver has error profinet network
      ER_U02_Servo_Fault : Bool;   // Servo driver has error
      WN_U02_Servo_Alarm : Bool;   // Servo driver has an warning
      ER_U02_Servo_STO_Active : Bool;   // Servo driver STO is active
      WN_U02_No_MemoryCard : Bool;   // Memory card is missing
      ER_U03_Servo_PN_NotPresent : Bool;   // Servo driver not present on profinet network
      ER_U03_Servo_PN_Error : Bool;   // Servo driver has error profinet network
      ER_U03_Servo_Fault : Bool;   // Servo driver has error
      WN_U03_Servo_Alarm : Bool;   // Servo driver has an warning
      ER_U03_Servo_STO_Active : Bool;   // Servo driver STO is active
      WN_U03_No_MemoryCard : Bool;   // Memory card is missing
      ER_U04_Servo_PN_NotPresent : Bool;   // Servo driver not present on profinet network
      ER_U04_Servo_PN_Error : Bool;   // Servo driver has error profinet network
      ER_U04_Servo_Fault : Bool;   // Servo driver has error
      WN_U04_Servo_Alarm : Bool;   // Servo driver has an warning
      ER_U04_Servo_STO_Active : Bool;   // Servo driver STO is active
      WN_U04_No_MemoryCard : Bool;   // Memory card is missing
      ER_U05_Servo_PN_NotPresent : Bool;   // Servo driver not present on profinet network
      ER_U05_Servo_PN_Error : Bool;   // Servo driver has error profinet network
      ER_U05_Servo_Fault : Bool;   // Servo driver has error
      WN_U05_Servo_Alarm : Bool;   // Servo driver has an warning
      ER_U05_Servo_STO_Active : Bool;   // Servo driver STO is active
      WN_U05_No_MemoryCard : Bool;   // Memory card is missing
      ER_U06_Servo_PN_NotPresent : Bool;   // Servo driver not present on profinet network
      ER_U06_Servo_PN_Error : Bool;   // Servo driver has error profinet network
      ER_U06_Servo_Fault : Bool;   // Servo driver has error
      WN_U06_Servo_Alarm : Bool;   // Servo driver has an warning
      ER_U06_Servo_STO_Active : Bool;   // Servo driver STO is active
      WN_U06_No_MemoryCard : Bool;   // Memory card is missing
      ER_U07_Servo_PN_NotPresent : Bool;   // Servo driver not present on profinet network
      ER_U07_Servo_PN_Error : Bool;   // Servo driver has error profinet network
      ER_U07_Servo_Fault : Bool;   // Servo driver has error
      WN_U07_Servo_Alarm : Bool;   // Servo driver has an warning
      ER_U07_Servo_STO_Active : Bool;   // Servo driver STO is active
      WN_U07_No_MemoryCard : Bool;   // Memory card is missing
      ER_U08_Servo_PN_NotPresent : Bool;   // Servo driver not present on profinet network
      ER_U08_Servo_PN_Error : Bool;   // Servo driver has error profinet network
      ER_U08_Servo_Fault : Bool;   // Servo driver has error
      WN_U08_Servo_Alarm : Bool;   // Servo driver has an warning
      ER_U08_Servo_STO_Active : Bool;   // Servo driver STO is active
      WN_U08_No_MemoryCard : Bool;   // Memory card is missing
      ER_U09_Servo_PN_NotPresent : Bool;   // Servo driver not present on profinet network
      ER_U09_Servo_PN_Error : Bool;   // Servo driver has error profinet network
      ER_U09_Servo_Fault : Bool;   // Servo driver has error
      WN_U09_Servo_Alarm : Bool;   // Servo driver has an warning
      ER_U09_Servo_STO_Active : Bool;   // Servo driver STO is active
      WN_U09_No_MemoryCard : Bool;   // Memory card is missing
      ER_U10_Servo_PN_NotPresent : Bool;   // Servo driver not present on profinet network
      ER_U10_Servo_PN_Error : Bool;   // Servo driver has error profinet network
      ER_U10_Servo_Fault : Bool;   // Servo driver has error
      WN_U10_Servo_Alarm : Bool;   // Servo driver has an warning
      ER_U10_Servo_STO_Active : Bool;   // Servo driver STO is active
      WN_U10_No_MemoryCard : Bool;   // Memory card is missing
      U01_FaultCode : Word;
      U01_AlarmCode : Word;
      U02_FaultCode : Word;
      U02_AlarmCode : Word;
      U03_FaultCode : Word;
      U03_AlarmCode : Word;
      U04_FaultCode : Word;
      U04_AlarmCode : Word;
      U05_FaultCode : Word;
      U05_AlarmCode : Word;
      U06_FaultCode : Word;
      U06_AlarmCode : Word;
      U07_FaultCode : Word;
      U07_AlarmCode : Word;
      U08_FaultCode : Word;
      U08_AlarmCode : Word;
      U09_FaultCode : Word;
      U09_AlarmCode : Word;
      U10_FaultCode : Word;
      U10_AlarmCode : Word;
   END_STRUCT;

END_TYPE

TYPE "UDT_MCC_IO"
TITLE = UDT_IO_MCC
VERSION : 0.1
//IO of main control cabinet
//# Block Info
//- Title:            UDT_IO_MCC
//- Comment/Function: IO of main control cabinet
//- Library/Family:   APS
//- Author:           Jay Liu
//- Tested with:      ---
//- Engineering:      TIA Portal V20
//- Restrictions:     ---
//- Requirements:     ---
//
//# History
// |Version  | Date       | Author                 | Description                   |
// |---------|------------|------------------------|------------------------------ |
// |01.00.00 | 2026-01-22 | Jay Liu                | First released version        |
   STRUCT
      Input : Struct
         Btn_Stop : Bool;
         Btn_Start : Bool;
         Btn_Reset : Bool;
         Cabinet_Temperature_High : Bool;
         PowerSupply_OK_G1011 : Bool;
         PowerSupply_OK_G1041 : Bool;
         Main_Switch_On_Q1001 : Bool;
         CB_F1011_On_Power_Supply : Bool;
         CB_F1012_On_UPS_Out : Bool;
         CB_F1021_On_HMI : Bool;
         CB_F1022_On_CPU : Bool;
         CB_F1023_On_XC216 : Bool;
         CB_F1024_On_Safety_XC208 : Bool;
         CB_F1025_On_Safety_CPU : Bool;
         CB_F1026_On_Image_Server : Bool;
         CB_F1031_On_Image_Switch : Bool;
         CB_F1032_On_HLC_Gateway : Bool;
         CB_F1033_On_Reserved : Bool;
         CB_F1034_On_Reserved : Bool;
         CB_F1072_On_PowerMeter_380VAC : Bool;
         CB_F1072_On_PowerMeter_220VAC : Bool;
         CB_F1041_On_Power_Supply : Bool;
         CB_F105x_On_GC03_Scanner : Bool;
         CB_F105x_On_GC04_Scanner : Bool;
         CB_F105x_On_Safety_IO_24VDC : Bool;
         CB_F105x_On_External_24VDC : Bool;
         CB_F1081_On_AC01 : Bool;
         CB_F1091_On_GC01_Inveter : Bool;
         CB_F1092_On_AC02 : Bool;
         CB_F1093_On_GC01_Interroll : Bool;
         CB_F1094_On_GC01_SDC01 : Bool;
         CB_F1101_On_GC02_Inveter : Bool;
         CB_F1102_On_AC03 : Bool;
         CB_F1103_On_Reversed : Bool;
         CB_F1104_On_GC02_SDC01 : Bool;
         CB_F1111_On_GC03_Inveter : Bool;
         CB_F1112_On_AC04 : Bool;
         CB_F1113_On_GC03_Interroll : Bool;
         CB_F1114_On_GC03_SDC01 : Bool;
         CB_F1115_On_GC03_SDC02 : Bool;
         CB_F1121_On_GC04_Inveter : Bool;
         CB_F1122_On_AC05 : Bool;
         CB_F1123_On_Reversed : Bool;
         CB_F1131_On_GC05_Inveter : Bool;
         CB_F1132_On_GC05_Interroll : Bool;
         CB_F1133_On_GC06_Inveter : Bool;
         CB_F1134_On_GC06_Interroll : Bool;
         CB_F1141_On_GC07_Inveter : Bool;
         CB_F1142_On_GC07_Interroll : Bool;
         CB_F1151_On_GC03_Inveter_Group2 : Bool;
         CB_F1152_On_Reversed : Bool;
         CB_F1153_On_Reversed : Bool;
         CB_F1154_On_Reversed : Bool;
         CB_F1155_On_EH01 : Bool;
         CB_F1156_On_EH02 : Bool;
         CB_F1157_On_EH03 : Bool;
         CB_F1161_On_Fan : Bool;
         CB_F1171_On_Socket : Bool;
         KM_1641_On_GC01_Interroll : Bool;
         KM_1642_On_GC01_Interroll : Bool;
         KM_1643_On_Reversed : Bool;
         KM_1644_On_Reversed : Bool;
         KM_1645_On_GC03_Interroll : Bool;
         KM_1646_On_GC03_Interroll : Bool;
         KM_1647_On_Reversed : Bool;
         KM_1648_On_Reversed : Bool;
         KM_1651_On_GC05_Interroll : Bool;
         KM_1652_On_GC05_Interroll : Bool;
         KM_1653_On_GC05_Interroll : Bool;
         KM_1654_On_GC05_Interroll : Bool;
         KM_1655_On_GC05_Interroll : Bool;
         KM_1656_On_GC05_Interroll : Bool;
      END_STRUCT;
      Output : Struct
         Light_Start_Btn : Bool;
         Light_Reset_Btn : Bool;
         Aux_On : Bool;
      END_STRUCT;
   END_STRUCT;

END_TYPE

TYPE "UDT_SDC_10Servos_IO"
VERSION : 0.1
   STRUCT
      Spare_0_0 : Bool;
      Spare_0_1 : Bool;
      Spare_0_2 : Bool;
      Spare_0_3 : Bool;
      Spare_0_4 : Bool;
      Spare_0_5 : Bool;
      Spare_0_6 : Bool;
      Spare_0_7 : Bool;
      Spare_1_0 : Bool;
      Spare_1_1 : Bool;
      Spare_1_2 : Bool;
      Spare_1_3 : Bool;
      Spare_1_4 : Bool;
      Spare_1_5 : Bool;
      Spare_1_6 : Bool;
      Spare_1_7 : Bool;
   END_STRUCT;

END_TYPE

TYPE "UDT_Tipper_Command"
VERSION : 0.1
   STRUCT
      Spare_0_0 : Bool;
      Spare_0_1 : Bool;
      Spare_0_2 : Bool;
      Spare_0_3 : Bool;
      Spare_0_4 : Bool;
      Spare_0_5 : Bool;
      Spare_0_6 : Bool;
      Spare_0_7 : Bool;
      Spare_1_0 : Bool;
      Spare_1_1 : Bool;
      Spare_1_2 : Bool;
      Spare_1_3 : Bool;
      Spare_1_4 : Bool;
      Spare_1_5 : Bool;
      Spare_1_6 : Bool;
      Spare_1_7 : Bool;
   END_STRUCT;

END_TYPE

FUNCTION_BLOCK "FB_Conv_MultiControl"
{ S7_Optimized_Access := 'TRUE' }
VERSION : 0.1
   VAR_INPUT
      i_IO_PEC_Position : Bool;
      i_IO_PEC_Trigger : Bool;
      i_Setting : "UDT_Conv_MultiControl_Setting";
      i_External_Request : "UDT_External_Request";
      i_Command : "UDT_Conv_MultiControl_Command";
   END_VAR

   VAR_OUTPUT RETAIN
      o_Status : "UDT_Conv_MultiControl_Status";
      o_General_Status : "UDT_General_Status";
      o_Diagnostics : "UDT_Conv_MultiControl_Diagnostics";
   END_VAR

   VAR_IN_OUT
      io_Global : "UDT_Global";
      io_System_Control : "UDT_System_Control";
      io_MultiControl_U01_IO : "UDT_MultiControl_HW_Interface";
      io_MultiControl_U02_IO : "UDT_MultiControl_HW_Interface";
      io_MultiControl_U03_IO : "UDT_MultiControl_HW_Interface";
      io_MultiControl_U04_IO : "UDT_MultiControl_HW_Interface";
      io_FIF_Upstream : "UDT_Flow_Interface";
      io_FIF : "UDT_Flow_Interface";
      io_FIF_Downstream : "UDT_Flow_Interface";
   END_VAR

   VAR
      s_FB_Displacement_AccDec : "FB_Displacement_AccDec";
      s_FB_EQP_PEC_Position : "FB_EQP_PEC_Position";
      s_FB_EQP_PEC_Trigger : "FB_EQP_PEC_Trigger";
      s_FB_EQP_Transport : "FB_EQP_Transport";
      s_FB_HW_MultiControl_U01 : "FB_HW_MultiControl";
      s_FB_HW_MultiControl_U02 : "FB_HW_MultiControl";
      s_FB_HW_MultiControl_U03 : "FB_HW_MultiControl";
      s_FB_HW_MultiControl_U04 : "FB_HW_MultiControl";
   END_VAR
   VAR RETAIN
      s_Cnt_PEC_Items { S7_SetPoint := 'True'} : Int;
      s_Speed_Select : Int;
      s_SW_Actual_Speed : Int;
      s_HW_U01_Actual_Speed : Int;
      s_HW_U02_Actual_Speed : Int;
      s_HW_U03_Actual_Speed : Int;
      s_HW_U04_Actual_Speed : Int;
      s_CMD_PEC_Preset_Latch : Bool;
      s_CMD_Motor : Bool;
      s_CMD_Motor_Reverse : Bool;
      s_HW_U01_Req_Halt : Bool;
      s_HW_U02_Req_Halt : Bool;
      s_HW_U03_Req_Halt : Bool;
      s_HW_U04_Req_Halt : Bool;
      s_PE_Position_Latch : Bool;
      s_PE_Trigger_Latch : Bool;
      s_Ext_Req_Stop : Bool;
      s_Ext_Req_Halt : Bool;
      s_Ext_Req_Disable_Send : Bool;
      s_Ext_Req_Disable_Recv : Bool;
      s_Ext_Req_Rest_ESave : Bool;
      s_Ext_Req_Clear_Data : Bool;
      s_SW_Motor_OnSpeed : Bool;
      s_HW_Motor_Running : Bool;
   END_VAR

   VAR_TEMP
      t_PEC_Position_Items : UDInt;
      t_PEC_Trigger_Items : UDInt;
      t_PEC_Position_Ready_To_Reset : Bool;
      t_PEC_Trigger_Ready_To_Reset : Bool;
      t_HW_VFD_U01_Ready_To_Reset : Bool;
      t_HW_VFD_U02_Ready_To_Reset : Bool;
      t_HW_VFD_U03_Ready_To_Reset : Bool;
      t_HW_VFD_U04_Ready_To_Reset : Bool;
      t_ER_Motor_U01_Fault : Bool;
      t_ER_Motor_U02_Fault : Bool;
      t_ER_Motor_U03_Fault : Bool;
      t_ER_Motor_U04_Fault : Bool;
      t_ER_Motor_Fault : Array[1..16] of Bool;
   END_VAR


BEGIN
	REGION NETWORK: Initial

	    FILL_BLK(IN    := FALSE,
	             COUNT := 16,
	             OUT   => #t_ER_Motor_Fault[1]);

	END_REGION

	REGION NETWORK AA: Conveyor Cycle Displacement
	    #s_FB_Displacement_AccDec(i_Conveyor_Speed   := #io_FIF.Speed,
	                              i_Accelaration     := #i_Setting.Hardware_U01.Acceleration,
	                              i_Decelaration     := #i_Setting.Hardware_U01.Deceleration,
	                              i_Prev_Cycle_Time  := #io_Global.OB_Prev_Cycle_Time,
	                              i_PPI_Displacement := 0,
	                              i_Section_Run      := #io_FIF.Motor_Run,
	                              o_Motor_On_Speed   => #o_General_Status.Motor_On_Speed,
	                              o_Motor_Stopped    => #io_FIF.Motor_Stopped,
	                              o_Actual_Speed     => #s_SW_Actual_Speed,
	                              o_Displacement     => #io_FIF.Displacement);

	    #o_General_Status.Motor_Stopped := #io_FIF.Motor_Stopped;
	END_REGION

	REGION NETWORK BA: Equipment layer - PEC
	    #s_FB_EQP_PEC_Position(i_IO_Available             := #io_System_Control.IO_Available,
	                           i_CMD_Reset                := #io_System_Control.OS_Reset_Jam,
	                           i_CMD_Clear_Stat           := #io_System_Control.OS_Clear_Statistics,
	                           i_CFG_Blockage_Length      := #i_Setting.PE1.Blockage_Length,
	                           i_CFG_Delay_On             := #i_Setting.PE1.Delay_On,
	                           i_CFG_Delay_Off            := #i_Setting.PE1.Delay_Off,
	                           i_CFG_Shifting_Offset      := #i_Setting.PE1.Shifting_Offset,
	                           i_CFG_Handover_Offset      := #i_Setting.PE1.Handover_Offset,
	                           i_CFG_Detect_PEC_OnStopped := #i_Setting.PE1.Detect_PEC_OnStopped,
	                           i_CFG_Reset_Block_PEC_Oc   := #i_Setting.PE1.Reset_Block_PEC_Oc,
	                           i_CFG_Item_On              := #i_Setting.PE1.Item_On,
	                           i_CMD_Preset_Latch         := #s_CMD_PEC_Preset_Latch,
	                           i_CMD_Clear_Data           := #s_Ext_Req_Clear_Data,
	                           i_Cycle_Count              := #io_FIF.Displacement,
	                           i_IO_PEC                   := #i_IO_PEC_Position,
	                           i_Section_Running          := NOT #io_FIF.Motor_Stopped,
	                           o_Ready_To_Reset           => #t_PEC_Position_Ready_To_Reset,
	                           o_ER_PEC_Blockage          => #o_Status.ER_PE1_Blockage,
	                           o_PEC_Filter               => #s_PE_Position_Latch,
	                           o_Handover                 => #io_FIF.Handover,
	                           o_Cnt_Buffer_Used          => #s_Cnt_PEC_Items,
	                           o_Stat_Items               => #t_PEC_Position_Items);

	    #s_FB_EQP_PEC_Trigger(i_IO_Available             := #io_System_Control.IO_Available,
	                          i_CMD_Reset                := #io_System_Control.OS_Reset_Jam,
	                          i_CMD_Clear_Stat           := #io_System_Control.OS_Clear_Statistics,
	                          i_CFG_Blockage_Length      := #i_Setting.PE2.Blockage_Length,
	                          i_CFG_Delay_On             := #i_Setting.PE2.Delay_On,
	                          i_CFG_Delay_Off            := #i_Setting.PE2.Delay_Off,
	                          i_CFG_Detect_PEC_OnStopped := #i_Setting.PE2.Detect_PEC_OnStopped,
	                          i_CFG_Reset_Block_PEC_Oc   := #i_Setting.PE2.Reset_Block_PEC_Oc,
	                          i_CFG_Item_On              := #i_Setting.PE2.Item_On,
	                          i_CMD_Preset_Latch         := false,
	                          i_Cycle_Count              := #io_FIF.Displacement,
	                          i_IO_PEC                   := #i_IO_PEC_Trigger,
	                          i_Section_Running          := NOT #io_FIF.Motor_Stopped,
	                          o_Ready_To_Reset           => #t_PEC_Trigger_Ready_To_Reset,
	                          o_ER_PEC_Blockage          => #o_Status.ER_PE2_Blockage,
	                          o_PEC_Filter               => #s_PE_Trigger_Latch,
	                          o_Stat_Items               => #t_PEC_Trigger_Items);

	    #io_FIF.PECTrigger_Latch := #s_PE_Trigger_Latch;
	END_REGION

	REGION NETWORK CA: Conditions to basic control
	    // Condition to request stop
	    #s_Ext_Req_Stop := #o_Status.ER_Motor_1_Fault
	    OR #o_Status.ER_Motor_2_Fault
	    OR #o_Status.ER_Motor_3_Fault
	    OR #o_Status.ER_Motor_4_Fault
	    OR #o_Status.ER_Motor_5_Fault
	    OR #o_Status.ER_Motor_6_Fault
	    OR #o_Status.ER_Motor_7_Fault
	    OR #o_Status.ER_Motor_8_Fault
	    OR #o_Status.ER_Motor_9_Fault
	    OR #o_Status.ER_Motor_10_Fault
	    OR #o_Status.ER_Motor_11_Fault
	    OR #o_Status.ER_Motor_12_Fault
	    OR #o_Status.ER_Motor_13_Fault
	    OR #o_Status.ER_Motor_14_Fault
	    OR #o_Status.ER_Motor_15_Fault
	    OR #o_Status.ER_Motor_16_Fault
	    OR #i_External_Request.Request_Stop;

	    // Condition to request halt
	    #s_Ext_Req_Halt := #s_HW_U01_Req_Halt
	    OR #s_HW_U02_Req_Halt
	    OR #s_HW_U03_Req_Halt
	    OR #s_HW_U04_Req_Halt
	    OR #i_External_Request.Request_Halt
	    OR #i_Command.Man_Mode
	    OR #o_Status.ER_PE1_Blockage
	    OR #o_Status.ER_PE2_Blockage;

